// ---- POUs/System/Functions/FindINTFieldFragmented.TcPOU
FUNCTION FindINTFieldFragmented : INT
VAR_INPUT
    FieldName : STRING(254);
    Str1 : STRING(254);
    Str2 : STRING(254);
END_VAR
VAR_OUTPUT
    Valid : BOOL;
END_VAR
VAR
    value : DINT;
END_VAR

FindINTFieldFragmented := -9999;
value := FindDINTFieldFragmented(FieldName := FieldName, Str1 := Str1, Str2 := Str2, Valid => Valid);
IF NOT Valid THEN RETURN; END_IF;
Valid := (value >= -32768) AND (value <= 32767);
IF Valid THEN FindINTFieldFragmented := DINT_TO_INT(value); END_IF;

END_FUNCTION

// ---- POUs/System/Functions/RemovePlusSign.TcPOU
FUNCTION RemovePlusSign : STRING(254)
VAR_INPUT
    inString : STRING(254);
END_VAR

// Preserve the reference behavior: remove only one leading plus sign.
RemovePlusSign := inString;
IF LEFT(inString, 1) = '+' THEN
    RemovePlusSign := RIGHT(inString, LEN(inString) - 1);
END_IF;

END_FUNCTION

// ---- POUs/System/Tests/FC_TestTIAFoundation.TcPOU
FUNCTION FC_TestTIAFoundation : DWORD
VAR
    value : WORD;
    success : BOOL;
    decoded : ID_Decoded_DUT;
    lamps : Stack_Lights_FB;
    result : STRING(254);
END_VAR

// Offline utility checks: return DWORD#0 when all checks pass.
// Invoke manually in an isolated test PLC. No physical I/O or global data is used.
// Failure bits identify the numbered checks below; no task call is installed.
FC_TestTIAFoundation := DWORD#0;

// Bit 0: set the highest WORD bit and preserve other bits.
value := WORD#16#0001;
success := Set_Bit_F(BIT_Number := 15, Bit_Value := TRUE, Variavel := value);
IF NOT success OR (value <> WORD#16#8001) THEN
    FC_TestTIAFoundation := FC_TestTIAFoundation OR DWORD#16#0001;
END_IF;
// Bit 1: FALSE is intentionally a no-op, not a reset operation.
success := Set_Bit_F(BIT_Number := 15, Bit_Value := FALSE, Variavel := value);
IF NOT success OR (value <> WORD#16#8001) THEN
    FC_TestTIAFoundation := FC_TestTIAFoundation OR DWORD#16#0002;
END_IF;
// Bit 2: reject out-of-range shifts without modifying the word.
success := Set_Bit_F(BIT_Number := 16, Bit_Value := TRUE, Variavel := value);
IF success OR (value <> WORD#16#8001) THEN
    FC_TestTIAFoundation := FC_TestTIAFoundation OR DWORD#16#0004;
END_IF;
// Bit 3: decimal ID decomposition.
success := ID_Decode_F(ID := 123456, ID_Decoded := decoded);
IF NOT success OR (decoded.Device_Type <> 12) OR
   (decoded.Level <> 34) OR (decoded.VTD <> 56) THEN
    FC_TestTIAFoundation := FC_TestTIAFoundation OR DWORD#16#0008;
END_IF;
// Bit 4: invalid ID must not retain the preceding decoded result.
success := ID_Decode_F(ID := -1, ID_Decoded := decoded);
IF success OR (decoded.Device_Type <> 0) OR (decoded.Level <> 0) OR (decoded.VTD <> 0) THEN
    FC_TestTIAFoundation := FC_TestTIAFoundation OR DWORD#16#0010;
END_IF;
// Bit 5: accept leading zero fields and the unassigned ID.
success := ID_Decode_F(ID := 0, ID_Decoded := decoded);
IF NOT success OR (decoded.Device_Type <> 0) OR (decoded.Level <> 0) OR (decoded.VTD <> 0) THEN
    FC_TestTIAFoundation := FC_TestTIAFoundation OR DWORD#16#0020;
END_IF;
// Bit 6: source-compatible SICK field spacing.
result := FindStringField(FieldName := 'Code', JsonStr := '{"Number" :"2", "Code" :"ABC123"}');
IF result <> 'ABC123' THEN
    FC_TestTIAFoundation := FC_TestTIAFoundation OR DWORD#16#0040;
END_IF;
// Bit 7: a barcode longer than the source's 10-character search window.
result := FindStringField(FieldName := 'Code', JsonStr := '{"Code":"123456789012345678901234567890"}');
IF result <> '123456789012345678901234567890' THEN
    FC_TestTIAFoundation := FC_TestTIAFoundation OR DWORD#16#0080;
END_IF;
// Bit 8: missing field returns empty after a previous successful call.
result := FindStringField(FieldName := 'Code', JsonStr := '{"Number":"3"}');
IF result <> '' THEN
    FC_TestTIAFoundation := FC_TestTIAFoundation OR DWORD#16#0100;
END_IF;
// Bit 9: an unterminated value must not be accepted.
result := FindStringField(FieldName := 'Code', JsonStr := '{"Code":"ABC');
IF result <> '' THEN
    FC_TestTIAFoundation := FC_TestTIAFoundation OR DWORD#16#0200;
END_IF;
// Bit 10: fault takes priority over automatic mode.
lamps(System_Auto := TRUE, Fault := TRUE, i_bFlash_05Hz := TRUE);
IF NOT lamps.Red OR lamps.Green OR lamps.Orange OR lamps.Yellow THEN
    FC_TestTIAFoundation := FC_TestTIAFoundation OR DWORD#16#0400;
END_IF;
// Bit 11: manual mode uses yellow/orange and clears red/green.
lamps(System_Auto := FALSE, Fault := FALSE, i_bFlash_05Hz := FALSE);
IF lamps.Red OR lamps.Green OR NOT lamps.Orange OR NOT lamps.Yellow THEN
    FC_TestTIAFoundation := FC_TestTIAFoundation OR DWORD#16#0800;
END_IF;
// Bit 12: upper ID boundary validation.
success := ID_Decode_F(ID := 1000000, ID_Decoded := decoded);
IF success OR (decoded.Device_Type <> 0) OR (decoded.Level <> 0) OR (decoded.VTD <> 0) THEN
    FC_TestTIAFoundation := FC_TestTIAFoundation OR DWORD#16#1000;
END_IF;

END_FUNCTION

// ---- POUs/System/Tests/FC_TestTIAParsing.TcPOU
FUNCTION FC_TestTIAParsing : DWORD
VAR
    valid : BOOL;
    booleanValue : BOOL;
    integerValue : INT;
    longValue : DINT;
    buffer : ARRAY[0..1024] OF BYTE;
    result : STRING(254);
    window1 : STRING(254);
    truncated : BOOL;
    i : INT;
END_VAR

// Run only in an isolated test PLC. Zero means all checks passed.
// Each set bit identifies the corresponding assertion below.
FC_TestTIAParsing := DWORD#0;
IF RemovePlusSign('+42') <> '42' THEN FC_TestTIAParsing := FC_TestTIAParsing OR SHL(DWORD#1, 0); END_IF;
IF RemovePlusSign('4+2') <> '4+2' THEN FC_TestTIAParsing := FC_TestTIAParsing OR SHL(DWORD#1, 1); END_IF;
booleanValue := FindBoolField(FieldName := 'x', JsonStr := '{"x": false, "y": true}', Valid => valid);
IF booleanValue OR NOT valid THEN FC_TestTIAParsing := FC_TestTIAParsing OR SHL(DWORD#1, 2); END_IF;
booleanValue := FindBoolField(FieldName := 'x', JsonStr := '{"y":true}', Valid => valid);
IF booleanValue OR valid THEN FC_TestTIAParsing := FC_TestTIAParsing OR SHL(DWORD#1, 3); END_IF;
booleanValue := FindBoolField(FieldName := 'x', JsonStr := '{"x" :$T true$R$N}', Valid => valid);
IF NOT booleanValue OR NOT valid THEN FC_TestTIAParsing := FC_TestTIAParsing OR SHL(DWORD#1, 4); END_IF;
integerValue := FindIntField(FieldName := 'x', JsonStr := '{"x":32767}', Valid => valid);
IF NOT valid OR (integerValue <> 32767) THEN FC_TestTIAParsing := FC_TestTIAParsing OR SHL(DWORD#1, 5); END_IF;
integerValue := FindIntField(FieldName := 'x', JsonStr := '{"x":-32768}', Valid => valid);
IF NOT valid OR (integerValue <> -32768) THEN FC_TestTIAParsing := FC_TestTIAParsing OR SHL(DWORD#1, 6); END_IF;
integerValue := FindIntField(FieldName := 'x', JsonStr := '{"x":32768}', Valid => valid);
IF valid OR (integerValue <> -9999) THEN FC_TestTIAParsing := FC_TestTIAParsing OR SHL(DWORD#1, 7); END_IF;
longValue := FindDINTFieldFragmented(FieldName := 'x', Str1 := '{"x":2147483647}', Str2 := '', Valid => valid);
IF NOT valid OR (longValue <> DINT#2147483647) THEN FC_TestTIAParsing := FC_TestTIAParsing OR SHL(DWORD#1, 8); END_IF;
longValue := FindDINTFieldFragmented(FieldName := 'x', Str1 := '{"x":-2147483648}', Str2 := '', Valid => valid);
IF NOT valid OR (longValue <> DINT#-2147483648) THEN FC_TestTIAParsing := FC_TestTIAParsing OR SHL(DWORD#1, 9); END_IF;
longValue := FindDINTFieldFragmented(FieldName := 'x', Str1 := '{"x":2147483648}', Str2 := '', Valid => valid);
IF valid OR (longValue <> -9999) THEN FC_TestTIAParsing := FC_TestTIAParsing OR SHL(DWORD#1, 10); END_IF;
integerValue := FindIntField(FieldName := 'x', JsonStr := '{"x":12.3}', Valid => valid);
IF valid THEN FC_TestTIAParsing := FC_TestTIAParsing OR SHL(DWORD#1, 11); END_IF;
integerValue := FindIntField(FieldName := 'x', JsonStr := '{"x":12', Valid => valid);
IF valid THEN FC_TestTIAParsing := FC_TestTIAParsing OR SHL(DWORD#1, 12); END_IF;
integerValue := FindIntField(FieldName := 'x', JsonStr := '{"x":-9999}', Valid => valid);
IF NOT valid OR (integerValue <> -9999) THEN FC_TestTIAParsing := FC_TestTIAParsing OR SHL(DWORD#1, 13); END_IF;
integerValue := FindINTFieldFragmented(FieldName := 'x', Str1 := 'partial', Str2 := ',"x":42}', Valid => valid);
IF NOT valid OR (integerValue <> 42) THEN FC_TestTIAParsing := FC_TestTIAParsing OR SHL(DWORD#1, 14); END_IF;
integerValue := FindINTFieldFragmented(FieldName := 'x', Str1 := '{"x":4', Str2 := '2}', Valid => valid);
IF valid THEN FC_TestTIAParsing := FC_TestTIAParsing OR SHL(DWORD#1, 15); END_IF;
FOR i := 0 TO 1024 DO buffer[i] := 0; END_FOR;
buffer[0] := 65; buffer[1] := 13; buffer[2] := 10; buffer[3] := 66;
result := ByteArrayToString(Lenght := 4, ByteArray := buffer, Truncated => truncated);
IF (result <> 'AB') OR truncated THEN FC_TestTIAParsing := FC_TestTIAParsing OR SHL(DWORD#1, 16); END_IF;
result := ByteArrayToString(Lenght := -1, ByteArray := buffer, Truncated => truncated);
IF (result <> '') OR NOT truncated THEN FC_TestTIAParsing := FC_TestTIAParsing OR SHL(DWORD#1, 17); END_IF;
FOR i := 0 TO 254 DO buffer[i] := 65; END_FOR;
result := ByteArrayToString(Lenght := 255, ByteArray := buffer, ByteArrayToString_1 => window1, Truncated => truncated);
IF (LEN(result) <> 254) OR (LEN(window1) <> 155) OR NOT truncated THEN FC_TestTIAParsing := FC_TestTIAParsing OR SHL(DWORD#1, 18); END_IF;
integerValue := FindIntField(FieldName := 'x', JsonStr := '{"x":01}', Valid => valid);
IF valid THEN FC_TestTIAParsing := FC_TestTIAParsing OR SHL(DWORD#1, 19); END_IF;

END_FUNCTION

// ---- POUs/VTD/Light_Bars_FB.TcPOU
FUNCTION_BLOCK Light_Bars_FB
VAR_INPUT
	VTD_Mode:  UINT;
	VTD_Speed:  INT;
	Fault:  BOOL;
	// Drive enable state of the VTD. Replaces the Siemens "SinaSpeed_VTD_DB_1".EnableAxis
	// (enable of the former G120 drive). Suggested source: VTD_Control.Motor.stStatus.bOutputStageEnabled (PI 1.2).
	i_bDriveEnabled:  BOOL;
END_VAR
VAR_OUTPUT
	Animation_B1:  BYTE;
	Color_B1:  BYTE;
	Speed_B1:  Byte;
	Animation_B2:  Byte;
	Color_B2:  Byte;
	Speed_B2:  BYTE;
END_VAR
VAR
END_VAR

//Commands for Light Bar

IF VTD_Mode = 0 AND NOT Fault THEN // (0)Disabled = No light  
    Animation_B1:= Animation_B2:= 0;
    
// SIEMENS-LEGACY: ELSIF VTD_Mode = 1 AND VTD_Speed = 0 AND  NOT Fault AND NOT "SinaSpeed_VTD_DB_1".EnableAxis THEN // (1)Manual= Yellow Stop
ELSIF VTD_Mode = 1 AND VTD_Speed = 0 AND  NOT Fault AND NOT i_bDriveEnabled THEN // (1)Manual= Yellow Stop
    Animation_B1 := Animation_B2 := 1;
    Color_B1 := Color_B2 := 4;
    
// SIEMENS-LEGACY: ELSIF VTD_Mode = 1 AND VTD_Speed > 0 AND VTD_Speed <= 33 AND  NOT Fault AND "SinaSpeed_VTD_DB_1".EnableAxis THEN // (1)Manual= Yellow until 33%
ELSIF VTD_Mode = 1 AND VTD_Speed > 0 AND VTD_Speed <= 33 AND  NOT Fault AND i_bDriveEnabled THEN // (1)Manual= Yellow until 33%
    Animation_B1 := Animation_B2 := 2;
    Speed_B1 := Speed_B2 := 2;
    Color_B1 := Color_B2 := 4;
    
ELSIF VTD_Mode = 1 AND VTD_Speed > 33 AND VTD_Speed <= 100 AND  NOT Fault THEN // (1)Manual= Yellow until 66%
    Animation_B1 := Animation_B2 := 2;
    Speed_B1 := Speed_B2 := 0;
    Color_B1 := Color_B2 := 4;
    
// ELSIF VTD_Mode = 1 AND VTD_Speed > 66 AND VTD_Speed <= 100 AND  NOT Fault THEN // (1)Manual= Yellow until 100%
//     Animation_B1 := Animation_B2 := 2;
//     Speed_B1 := Speed_B2 := 1;
//     Color_B1 := Color_B2 := 4;
    
// SIEMENS-LEGACY: ELSIF VTD_Mode = 2 AND VTD_Speed = 0 AND  NOT Fault AND NOT "SinaSpeed_VTD_DB_1".EnableAxis THEN // (2)Semi-auto = Blue Stop
ELSIF VTD_Mode = 2 AND VTD_Speed = 0 AND  NOT Fault AND NOT i_bDriveEnabled THEN // (2)Semi-auto = Blue Stop
    Animation_B1 := Animation_B2 := 1;
    Color_B1 := Color_B2 := 9;
    Speed_B1 := Speed_B2 := 0;
    
// SIEMENS-LEGACY: ELSIF VTD_Mode = 2 AND VTD_Speed > 0 AND VTD_Speed <= 33 AND  NOT Fault AND "SinaSpeed_VTD_DB_1".EnableAxis THEN // (2)Semi-auto = Blue until 33%
ELSIF VTD_Mode = 2 AND VTD_Speed > 0 AND VTD_Speed <= 33 AND  NOT Fault AND i_bDriveEnabled THEN // (2)Semi-auto = Blue until 33%
    Animation_B1 := Animation_B2 := 2;
    Speed_B1 := Speed_B2 := 2;
    Color_B1 := Color_B2 := 9;
    
ELSIF VTD_Mode = 2 AND VTD_Speed > 33 AND VTD_Speed <= 100 AND  NOT Fault THEN // (2)Semi-auto = Blue until 66%
    Animation_B1 := Animation_B2 := 2;
    Speed_B1 := Speed_B2 := 0;
    Color_B1 := Color_B2 := 9;
    
// ELSIF VTD_Mode = 2 AND VTD_Speed > 66 AND VTD_Speed <= 100 AND  NOT Fault THEN // (2)Semi-auto = Blue until 100%
//     Animation_B1 := Animation_B2 := 2;
//     Speed_B1 := Speed_B2 := 1;
//     Color_B1 := Color_B2 := 9;
    
// SIEMENS-LEGACY: ELSIF VTD_Mode = 3 AND VTD_Speed = 0 AND  NOT Fault AND NOT "SinaSpeed_VTD_DB_1".EnableAxis THEN // (3)Auto = Green Stop
ELSIF VTD_Mode = 3 AND VTD_Speed = 0 AND  NOT Fault AND NOT i_bDriveEnabled THEN // (3)Auto = Green Stop
    Animation_B1 := Animation_B2 := 1;
    Color_B1 := Color_B2 := 0;
    
// SIEMENS-LEGACY: ELSIF VTD_Mode = 3 AND VTD_Speed > 0 AND VTD_Speed <= 33 AND  NOT Fault AND "SinaSpeed_VTD_DB_1".EnableAxis THEN // (3)Auto = Green until 33%
ELSIF VTD_Mode = 3 AND VTD_Speed > 0 AND VTD_Speed <= 33 AND  NOT Fault AND i_bDriveEnabled THEN // (3)Auto = Green until 33%
    Animation_B1 := Animation_B2 := 2;
    Speed_B1 := Speed_B2 := 2;
    Color_B1 := Color_B2 := 0;
    
ELSIF VTD_Mode = 3 AND VTD_Speed > 33 AND VTD_Speed <= 100 AND  NOT Fault THEN // (3)Auto = Green until 66%
    Animation_B1 := Animation_B2 := 2;
    Speed_B1 := Speed_B2 := 0;
    Color_B1 := Color_B2 := 0;
    
// ELSIF VTD_Mode = 3 AND VTD_Speed > 66 AND VTD_Speed <= 100 AND  NOT Fault THEN // (3)Auto = Green until 100%
//     Animation_B1 := Animation_B2 := 2;
//     Speed_B1 := Speed_B2 := 1;
//     Color_B1 := Color_B2 := 0;
    
ELSIF VTD_Mode = 4 AND VTD_Speed = 0 AND  NOT Fault THEN // (4)Tech = Orange Stop
    Animation_B1 := Animation_B2 := 1;
    Color_B1 := Color_B2 := 2;
    
ELSIF VTD_Mode = 4 AND VTD_Speed > 0 AND VTD_Speed <= 33 AND  NOT Fault THEN // (4)Tech = Orange until 33%
    Animation_B1 := Animation_B2 := 2;
    Speed_B1 := Speed_B2 := 2;
    Color_B1 := Color_B2 := 2;
    
ELSIF VTD_Mode = 4 AND VTD_Speed > 33 AND VTD_Speed <= 66 AND  NOT Fault THEN // (4)Tech = Orange until 66%
    Animation_B1 := Animation_B2 := 2;
    Speed_B1 := Speed_B2 := 0;
    Color_B1 := Color_B2 := 2;
    
ELSIF VTD_Mode = 4 AND VTD_Speed > 66 AND VTD_Speed <= 100 AND  NOT Fault THEN // (4)Tech = Orange until 100%
    Animation_B1 := Animation_B2 := 2;
    Speed_B1 := Speed_B2 := 1;
    Color_B1 := Color_B2 := 2;
    
ELSIF VTD_Mode = 5 AND VTD_Speed = 0 AND  NOT Fault THEN // (5)Maintenance = White Stop
    Animation_B1 := Animation_B2 := 1;
    Color_B1 := Color_B2 := 19;
    
ELSIF VTD_Mode = 5 AND VTD_Speed > 0 AND VTD_Speed <= 33 AND  NOT Fault THEN // (5)Maintenance = White until 33%
    Animation_B1 := Animation_B2 := 2;
    Speed_B1 := Speed_B2 := 2;
    Color_B1 := Color_B2 := 19;
    
ELSIF VTD_Mode = 5 AND VTD_Speed > 33 AND VTD_Speed <= 66 AND  NOT Fault THEN // (5)Maintenance = White until 66%
    Animation_B1 := Animation_B2 := 2;
    Speed_B1 := Speed_B2 := 0;
    Color_B1 := Color_B2 := 19;
    
ELSIF VTD_Mode = 5 AND VTD_Speed > 66 AND VTD_Speed <= 100 AND  NOT Fault THEN // (5)Maintenance = White until 100%
    Animation_B1 := Animation_B2 := 2;
    Speed_B1 := Speed_B2 := 1;
    Color_B1 := Color_B2 := 19;
    
ELSIF Fault THEN // Fault = Flash Red
    Animation_B1:= Animation_B2 := 2;
    Color_B1:=Color_B2 := 1;
END_IF;

END_FUNCTION_BLOCK

// ---- POUs/VTD/VTD_FB.TcPOU
FUNCTION_BLOCK VTD_FB
VAR_INPUT
	System_no:  UINT;
	Safety_OK:  BOOL;
	Cnv_Sensors:  Cnv_Inputs_DUT;
	VTD_Settings:  VTD_Settings_DUT;
	Bypass_DP:  BOOL;
// 	Bypass:  Safety_Bypass_RemotePanel;
END_VAR
VAR_OUTPUT
END_VAR
VAR_IN_OUT
	VTD_Control:  VTD_Control_DUT;
	LE_Bypass_HMI:  BOOL;
END_VAR
VAR
	State:  UINT;
	Last_State:  UINT;
	I_State:  UInt;
	LD_Timer_1:  TON;
	LD_Timer:  TON;
	DP_Timer:  TON;
	Watchdog:  TON;
	CS_TImer:  TON;
	Interlock_Timer:  TON;
	MainSetpoint:  Int;
	Position_Offset:  Real;
	ChangeToLow:  Array[1..4] of DInt;
	DestPosition:  Real;
	SetUpSpeed:  UInt;
	LevelBelowExtractor:  UInt;
	IEC_Timer_0_Instance:  TON;
	DestinationLevel:  UInt;
	CurrentlLevel:  UInt;
	VTD_ID_Decoded:  ID_Decoded_DUT;
	Cnv_ID_Decoded:  ARRAY[1..2] OF ID_Decoded_DUT;
	IEC_Timer_0_Instance_1:  TON;
	IEC_Timer_0_Instance_2:  TON;
	VTD_ControlInstructionTask_ID_Old:  Int;
	R_Execulte:  R_TRIG;
	R_AutomatcMode:  R_TRIG;
	T_Encoders_Difference:  TON;
	T_LE_Error:  TON;
	T_Setpoint_Delay:  TON;
	Distance_mm:  Real;
	TravelTime_s:  UInt;
	LE_Prev_mm:  Real;
	DeltaPos_mm:  Real;
	SampleTime_s:  Real;
	VTDSpeed_mm_s:  Real;
	T_Speed:  TON;
	Speed_mm_per_percent:  Real;
	Speed_mm_s:  Real;
	TravelTime_ms:  UInt;
	Watchdog_PT:  Time;
	Position_OLD:  Real;
	R_Position_OLD:  R_TRIG;

	// VTD drive: SEW MOVIPRO, MOVIKIT Positioning Drive (region "VFD")
	fbSewDrive:  FB_SEW_Drive;
	bDriveMoveRequest:  BOOL;
	bDriveEnable:  BOOL;
	bDriveFaultReset:  BOOL;
	rSpeedSetpoint:  REAL;              // [user units], signed
	rAccelerationFactor_pct:  REAL;     // [%] of SEW_Ramp_At_100pct
	uiDriveRamp:  UINT;                 // [user units]
	diPalletWeight:  DINT;
END_VAR

VAR_TEMP
	Level_Accuracy:  STRING;
	i:  UINT;
	Upper_limit:  Bool;
	Ultimate_SlowDown:  Bool;
	Ultimate_Creep:  Bool;
	Lower_Limit:  Bool;
	Level_Detect:  Bool;
	Level_Detect1:  Bool;
	Level_Detect2:  Bool;
	DP2_Extended:  Bool;
	DP2_Retracted:  Bool;
	DP1_Extended:  Bool;
	DP1_Retracted:  Bool;
	Chain_Slack_1:  Bool;
	Chain_Slack_2:  Bool;
	Chain_Slack_3:  Bool;
	Chain_Slack_4:  Bool;
	DP1_Retract:  Bool;
	DP1_Extend:  Bool;
	DP2_Retract:  Bool;
	DP2_Extend:  Bool;
	Cnvs1_NotExtended:  Bool;
	Cnvs2_NotExtended:  Bool;
	Stoppers_NotExtended:  Bool;
	MainSetpoint1:  Int;
	HMI_Reset:  BOOL;
END_VAR

// //Execute
// R_Execulte(CLK := VTD_Control.Instruction.Execulte);
// 
// IF VTD_Control.Mode = 3 THEN
//     VTD_Control.Instruction.Enable := TRUE;
// END_IF;
// 
// VTD_Control.Enabled := VTD_Control.Instruction.Enable;
// 
// VTD_Control.Mode := VTD_Control.Instruction.Mode_Change;
// 
// IF NOT VTD_Control.Enabled AND NOT VTD_Control.Error THEN
//     State := 0;
// END_IF;
// 
// //MANUAL MODE
// IF (VTD_Control.Mode = 1 OR VTD_Control.Mode = 5) AND NOT VTD_Control.Error AND VTD_Control.Enabled THEN
//     State := 500;
// END_IF;
// 
// (*
// TODO:
// 
// Mode select is done via the HMI. Might add external mode select switches.
//         
//         Mode select mask:
//         0: Disabled
//         1: Manual
//         2: Semi-Auto
//         3: Auto
//         4: Teach
//         5: Maintenance
//         
// Device ID Format: XXYYZZ    
// XX = Device type   
//     01   VTD
//     10  Cnv_Front_of_VTD
//     11  Cnv_Rear_of_VTD
//     12  Cnv_On_Extractor
//     20  Safety_Stop_Front_of_VTD
//     21  Safety_Stop_Rear_of_VTD
// YY = Floor   
// ZZ = VTD Connected to 
// *)
// 
// {region "Sensor allocations"}
//     //Assign inputs to local vars
//     Upper_limit := VTD_Control.Inputs.Upper_limit;
//     Ultimate_SlowDown := VTD_Control.Inputs.Ultimate_SlowDown;
//     Ultimate_Creep := VTD_Control.Inputs.Ultimate_Creep;
//     Lower_Limit := VTD_Control.Inputs.Lower_Limit;
//     Level_Detect1 := VTD_Control.Inputs.Level_Detect1;
//     Level_Detect2 := VTD_Control.Inputs.Level_Detect2;
//     DP1_Extended := VTD_Control.Inputs.DP1_Extended;
//     DP1_Retracted := VTD_Control.Inputs.DP1_Retracted;
//     DP2_Extended := VTD_Control.Inputs.DP2_Extended;
//     DP2_Retracted := VTD_Control.Inputs.DP2_Retracted;
//     Chain_Slack_1 := VTD_Control.Inputs.Chain_Slack_1;
//     Chain_Slack_2 := VTD_Control.Inputs.Chain_Slack_2;
//     Chain_Slack_3 := VTD_Control.Inputs.Chain_Slack_3;
//     Chain_Slack_4 := VTD_Control.Inputs.Chain_Slack_4;
//     VTD_Control.LinearEnc := VTD_Control.Inputs.LE_Position;
//     VTD_Control.AE := VTD_Control.Inputs.AE_Position_1;
// {endregion}
// 
// {region "Cyclic Checks"}
//     // Check for Pallet
//     IF Cnv_Sensors.Forward_Sensor OR Cnv_Sensors.Backward_Sensor THEN
//         VTD_Control.Pallet_Loaded := 1;//'Unknown';
//     ELSE
//         //No Pallet
//         VTD_Control.Pallet_Loaded := 0;//'None';
//     END_IF;
//     
//     //Docking pins
//         IF DP1_Extended AND DP2_Extended THEN
//             VTD_Control.LP_State := 1; //'Extended'
//         ELSIF DP1_Retracted AND DP2_Retracted THEN
//             VTD_Control.LP_State := 2; //'Retracted'
//         ELSE
//             VTD_Control.LP_State := 0; //'Unknown'
//         END_IF;
//         
//         VTD_Control.DP_Extended := VTD_Control.LP_State = 1;
//     
//     // Level detect
//     Level_Detect := Level_Detect1 AND Level_Detect2;
//     
//     //VTD extractor is docked
//     IF DP1_Extended AND DP2_Extended AND Level_Detect AND
//         (VTD_Control.LinearEnc - VTD_Settings.Teach_Values.Levels_LE[LevelBelowExtractor]) <= VTD_Settings.Level_Detect_LE THEN
//         VTD_Control.Docked := TRUE;
//     ELSE
//         VTD_Control.Docked := FALSE;
//     END_IF;
//     
//     //Ultimate stop checks
//     IF (VTD_Control.LinearEnc < VTD_Settings.Slowdown_Count_LE OR VTD_Control.LinearEnc > VTD_Settings.Teach_Values.Levels_LE[VTD_Settings.Highest_Level] - VTD_Settings.Slowdown_Count_LE) AND
//         Ultimate_Creep AND Ultimate_SlowDown AND VTD_Control.Running THEN
//         VTD_Control.Motor_Speed := VTD_Settings.Creep_Speed;
//         VTD_Control.Warning := 3; // Overtravel creep zone reached
//     ELSIF (VTD_Control.LinearEnc < VTD_Settings.Slowdown_Count_LE OR VTD_Control.LinearEnc > VTD_Settings.Teach_Values.Levels_LE[VTD_Settings.Highest_Level] - VTD_Settings.Slowdown_Count_LE) AND
//         NOT Ultimate_Creep AND Ultimate_SlowDown AND VTD_Control.Running THEN
//         VTD_Control.Motor_Speed := VTD_Settings.Slow_Speed; // Overtravel slow zone reached
//     END_IF;
//     
//     //Update Variables
//     IF VTD_Control.Current_Task_Type = 0 OR VTD_Control.Current_Task_Type = 1 THEN
//         VTD_Control.SM_State := State;
//     ELSIF VTD_Control.Current_Task_Type = 2 OR VTD_Control.Current_Task_Type = 3 THEN
//         VTD_Control.SM_State := I_State;
//     END_IF;
//     
//     FOR i := VTD_Settings.Lowest_Level TO VTD_Settings.Highest_Level DO
//         IF NOT Control.LCnv_Sys[System_no].Cnv_Level[i].Cnv1.Safety_Stop_Cnrl.Inputs.DP_Extended THEN
//             Cnvs1_NotExtended := true;
//         END_IF;
//         IF NOT Control.LCnv_Sys[System_no].Cnv_Level[i].Cnv2.Safety_Stop_Cnrl.Inputs.DP_Extended THEN
//             Cnvs2_NotExtended := true;
//         END_IF;
//     END_FOR;
//     
//     //Confirm whish level is below the extractor
//     FOR i := VTD_Settings.Lowest_Level TO VTD_Settings.Highest_Level DO
//         IF VTD_Control.LinearEnc >= (VTD_Settings.Teach_Values.Levels_LE[i] - VTD_Settings.Level_Detect_LE) THEN
//             LevelBelowExtractor := i;
//         END_IF;
//     END_FOR;
//     
//     Stoppers_NotExtended := Cnvs1_NotExtended (*AND Cnvs2_NotExtended*);
//     
//     //AE ERROR
//     IF VTD_Control.Inputs.AE_Status_2.15 THEN
//         VTD_Control.AE_Error := 1;
//     ELSE
//         VTD_Control.AE_Error := 0;
//     END_IF;
//     
//     //Encoder Delta
//     VTD_Control.Encoder_Delta := ABS(VTD_Control.AE - VTD_Control.LinearEnc);
//     
//     //CURRENT LEVEL
//     FOR i := VTD_Settings.Lowest_Level TO VTD_Settings.Highest_Level DO
//         IF ABS(VTD_Control.LinearEnc - VTD_Settings.Teach_Values.Levels_LE[i]) <= VTD_Settings.VTD_Level_Granularity AND Level_Detect THEN
//             VTD_Control.Current_Level := i;
//             EXIT;
//         ELSE
//             VTD_Control.Current_Level := 0;
//         END_IF;
//     END_FOR;
//     
//     //SPEED mm/S
//     T_Speed(IN := TRUE,
//              PT := T#100MS);
//     
//     IF T_Speed.Q THEN
//         DeltaPos_mm := ABS(VTD_Control.LinearEnc - LE_Prev_mm);
//         VTDSpeed_mm_s := DeltaPos_mm / SampleTime_s;
//         LE_Prev_mm := VTD_Control.LinearEnc;
//         T_Speed(IN := FALSE,
//                  PT := T#0MS);
//     END_IF;
// {endregion}
// 
// {region "Auto/Semi-Auto Mode"}
//     CASE State OF
//         0: //Idle
//             Last_State := State;
//             VTD_Control.Motor_UP := FALSE;
//             VTD_Control.Motor_Down := FALSE;
//             VTD_Control.Motor_Speed := 0; // SEW: was Motor.Speed
//             DestinationLevel := CurrentlLevel := 0;
//             VTD_Control.Stopped := TRUE;
//             Watchdog(IN := FALSE,
//                           PT := T#0S);
//             IF VTD_Control.Mode = 3 OR VTD_Control.Mode = 2 THEN
//                 IF VTD_Control.Instruction.Enable AND NOT VTD_Control.Error THEN
//                     State := 10;
//                 END_IF;
//             END_IF;
//             
//         10: //Standby
//             Last_State := State;
//             IF VTD_Control.Enabled AND NOT VTD_Control.Running AND VTD_Control.Instruction.Move_To_Level >= VTD_Settings.Lowest_Level AND
//                 VTD_Control.Instruction.Move_To_Level <= VTD_Settings.Highest_Level AND VTD_Control.Pallet_Loaded <> 1 AND
//                 ((VTD_Control.Instruction.Task_ID > 0 OR VTD_Control.Instruction.Task_Metadata <> '' AND VTD_Control.Mode = 3 AND Control.VTD_Order_Table[System_no].Task_Type = 1) OR
//                 (VTD_Control.Mode = 2 (*AND R_Execulte.Q*)))
//             THEN
//                 IF VTD_Control.Instruction.Move_To_Level = VTD_Control.Current_Level AND VTD_Control.Instruction.Move_To_Level <> 0 THEN
//                     VTD_Control.Warning := 1; //VTD already at level requested
//                     VTD_Control.Instruction.Move_To_Level := 0;
//                     //Go straght to the travel complete feedabck 
//                 ELSIF ((VTD_Control.Shuttle_Loaded = 0 OR VTD_Control.Shuttle_Loaded = 1) AND System_no <= 3)
//                     OR System_no > 3
//                 THEN //EVERYTHING OK
//                     DestinationLevel := VTD_Control.Instruction.Move_To_Level;
//                     CurrentlLevel := VTD_Control.Current_Level;
//                     VTD_Control.Current_Task_ID := VTD_Control.Instruction.Task_ID;
//                     VTD_Control.Running := TRUE;
//                     State := 20;
//                 END_IF;
//             END_IF;
// 
//         20: //Extend all safety stoppers that are not in the up position
//             Last_State := State;
//             VTD_Control.Done := FALSE;// To report to order table
//             FOR i := VTD_Settings.Lowest_Level TO VTD_Settings.Highest_Level DO
//                 IF NOT Control.LCnv_Sys[System_no].Cnv_Level[i].Cnv1.Safety_Stop_Cnrl.Inputs.DP_Extended THEN
//                     Control.LCnv_Sys[System_no].Cnv_Level[i].Cnv1.Safety_Stop_Cnrl.Instruction.Extend := TRUE;
//                 END_IF;
//                 IF NOT Control.LCnv_Sys[System_no].Cnv_Level[i].Cnv2.Safety_Stop_Cnrl.Inputs.DP_Extended THEN
//                     Control.LCnv_Sys[System_no].Cnv_Level[i].Cnv2.Safety_Stop_Cnrl.Instruction.Extend := TRUE;
//                 END_IF;
//             END_FOR;
//             State := 25;
//             
//         25: //Check to ensure the Safety stoppers are in the up position.
//             Last_State := State;
//             FOR i := VTD_Settings.Lowest_Level TO VTD_Settings.Highest_Level DO
//                 IF Control.LCnv_Sys[System_no].Cnv_Level[i].Cnv1.Safety_Stop_Cnrl.Inputs.DP_Extended THEN
//                     Control.LCnv_Sys[System_no].Cnv_Level[i].Cnv1.Safety_Stop_Cnrl.Instruction.Extend := FALSE;
//                 END_IF;
//                 IF Control.LCnv_Sys[System_no].Cnv_Level[i].Cnv2.Safety_Stop_Cnrl.Inputs.DP_Extended THEN
//                     Control.LCnv_Sys[System_no].Cnv_Level[i].Cnv2.Safety_Stop_Cnrl.Instruction.Extend := FALSE;
//                 END_IF;
//             END_FOR;
//             
//             IF Control.LCnv_Sys[System_no].Cnv_Level[2].Cnv1.Safety_Stop_Cnrl.Inputs.DP_Extended AND
//                 Control.LCnv_Sys[System_no].Cnv_Level[3].Cnv1.Safety_Stop_Cnrl.Inputs.DP_Extended AND
//                 Control.LCnv_Sys[System_no].Cnv_Level[4].Cnv1.Safety_Stop_Cnrl.Inputs.DP_Extended AND
//                 Control.LCnv_Sys[System_no].Cnv_Level[5].Cnv1.Safety_Stop_Cnrl.Inputs.DP_Extended AND
//                 Control.LCnv_Sys[System_no].Cnv_Level[6].Cnv1.Safety_Stop_Cnrl.Inputs.DP_Extended AND
//                 Control.LCnv_Sys[System_no].Cnv_Level[2].Cnv2.Safety_Stop_Cnrl.Inputs.DP_Extended AND
//                 Control.LCnv_Sys[System_no].Cnv_Level[3].Cnv2.Safety_Stop_Cnrl.Inputs.DP_Extended AND
//                 Control.LCnv_Sys[System_no].Cnv_Level[4].Cnv2.Safety_Stop_Cnrl.Inputs.DP_Extended AND
//                 Control.LCnv_Sys[System_no].Cnv_Level[5].Cnv2.Safety_Stop_Cnrl.Inputs.DP_Extended AND
//                 Control.LCnv_Sys[System_no].Cnv_Level[6].Cnv2.Safety_Stop_Cnrl.Inputs.DP_Extended
//             THEN
//                 State := 30;
//             END_IF;
//             
//         30: //Undock the VTD
//             Last_State := State;
//             IF LevelBelowExtractor >= VTD_Settings.Lowest_Level AND LevelBelowExtractor < VTD_Settings.Highest_Level THEN
//                 IF VTD_Control.Docked OR
//                     (VTD_Control.LinearEnc < VTD_Settings.Teach_Values.Levels_LE[LevelBelowExtractor] + 50) OR
//                     (VTD_Control.LinearEnc < VTD_Settings.Teach_Values.Levels_LE[LevelBelowExtractor + 1] AND
//                     VTD_Control.LinearEnc > VTD_Settings.Teach_Values.Levels_LE[LevelBelowExtractor + 1] - 10) THEN
//                     IF VTD_Control.LP_State = 1 THEN //extended
//                         VTD_Control.Motor_Speed := VTD_Settings.Dock_speed;
//                         VTD_Control.Motor_UP := TRUE;
//                         Position_Offset := VTD_Control.LinearEnc + 40;
//                         State := 35;
//                     ELSIF VTD_Control.LP_State = 2 THEN //retracted
//                         State := 45;
//                     ELSE //24:4 Docking pins in an known state
//                         Set_Bit_F(Bit_Number := 5,
//                                     Bit_Value := 1,
//                                     Variavel := VTD_Control.VTD_Errors.Error_Word_2);
//                     END_IF;
//                 ELSE
//                     Position_Offset := VTD_Control.LinearEnc - 5;
//                     State := 35;
//                 END_IF;
//             ELSIF LevelBelowExtractor = VTD_Settings.Highest_Level THEN
//                 IF VTD_Control.Docked OR
//                     (VTD_Control.LinearEnc < VTD_Settings.Teach_Values.Levels_LE[LevelBelowExtractor] + 50) THEN
//                     IF VTD_Control.LP_State = 1 THEN //extended
//                         VTD_Control.Motor_Speed := VTD_Settings.Dock_speed;
//                         VTD_Control.Motor_UP := TRUE;
//                         Position_Offset := VTD_Control.LinearEnc + 40;
//                         State := 35;
//                     ELSIF VTD_Control.LP_State = 2 THEN //retracted
//                         State := 45;
//                     ELSE //24:4 Docking pins in an known state
//                         Set_Bit_F(Bit_Number := 5,
//                                     Variavel := VTD_Control.VTD_Errors.Error_Word_2);
//                     END_IF;
//                 ELSE
//                     Position_Offset := VTD_Control.LinearEnc - 5;
//                     State := 35;
//                 END_IF;
//             END_IF;
//             
//         35: //Stop motor
//             Last_State := State;
//             IF NOT Level_Detect AND VTD_Control.LinearEnc >= Position_Offset THEN
//                 VTD_Control.Motor_Speed := 0;
//                 VTD_Control.Motor_UP := FALSE;
//                 State := 36;
//             END_IF;
//             
//         36: //Retract the docking pins
//             Last_State := State;
//                 DP2_Retract := DP1_Retract := TRUE;
//                 DP_Timer(IN := TRUE,
//                           PT := UINT_TO_TIME(VTD_Settings.Lockpins_Timeout_Retract));
//                 
//                 IF DP2_Retracted THEN
//                     DP2_Retract := FALSE;
//                 END_IF;
//                 IF VTD_Control.Inputs.DP1_Retracted THEN
//                     DP1_Retract := FALSE;
//                 END_IF;
//                 
//                 IF VTD_Control.LP_State = 2 THEN
//                     State := 40;
//                 END_IF;
//                 
//             40: //Check docking pins have been retracted
//                 Last_State := State;
//             IF VTD_Control.LP_State = 2 THEN
//                 DP_Timer(IN := FALSE,
//                           PT := T#0S);
//                 DP2_Retract := DP1_Retract := FALSE;
//                 State := 45;
//             END_IF;
//             
//         45: //Start moving towards the level required
//             Last_State := State;
//             //Check load type and set extractor speed
//             IF VTD_Control.Shuttle_Loaded = 0 AND VTD_Control.Pallet_Loaded = 0 THEN
//                 VTD_Control.Motor_Speed := VTD_Settings.Empty_Speed;
//             ELSIF VTD_Control.Shuttle_Loaded = 1 AND VTD_Control.Pallet_Loaded = 0 THEN
//                 VTD_Control.Motor_Speed := VTD_Settings.Shuttle_Speed;
//             ELSIF VTD_Control.Shuttle_Loaded = 0 AND (VTD_Control.Pallet_Loaded > 0) THEN
//                 VTD_Control.Motor_Speed := VTD_Settings.Pallet_Speed;
//             ELSIF VTD_Control.Shuttle_Loaded = 1 AND (VTD_Control.Pallet_Loaded > 0) THEN
//                 VTD_Control.Motor_Speed := VTD_Settings.Loaded_Speed;
//             END_IF;
//             
//             DestPosition := VTD_Settings.Teach_Values.Levels_LE[VTD_Control.Instruction.Move_To_Level];
//             SetUpSpeed := VTD_Control.Motor_Speed;
//             
//             // === DINAMIC WATCHDOG ===
//             Speed_mm_s := SetUpSpeed * Speed_mm_per_percent;
//             Distance_mm := ABS(DestPosition - VTD_Control.LinearEnc);
//             
//             //VTD needs to move up
//             IF VTD_Control.LinearEnc < DestPosition THEN
//                 VTD_Control.Motor_UP := TRUE;
//                 State := 50;
//                 //VTD needs to move down
//             ELSIF VTD_Control.LinearEnc > DestPosition THEN
//                 VTD_Control.Motor_Down := TRUE;
//                 State := 65; //change to 65
//             END_IF;
//             
//         50: //travel upwards to designated level
//             Last_State := State;
//             ChangeToLow[1] := ABS((VTD_Settings.Slowdown_Count_LE / 100) * 80); (* 80% *) //80  600mm
//             ChangeToLow[2] := ABS((VTD_Settings.Slowdown_Count_LE / 100) * 60); (* 60% *) //60
//             ChangeToLow[3] := ABS((VTD_Settings.Slowdown_Count_LE / 100) * 40); (* 40% *) //40
//             ChangeToLow[4] := ABS((VTD_Settings.Slowdown_Count_LE / 100) * 20); (* 20% *) //20 60
//             
//             //switch to fast freq Low UP
//             IF ABS(DestPosition - VTD_Control.LinearEnc) > VTD_Settings.Slowdown_Count_LE THEN
//                 VTD_Control.Motor_Speed := SetUpSpeed; //5
//                 //switch to low freq
//             ELSIF ABS(DestPosition - VTD_Control.LinearEnc) <= VTD_Settings.Slowdown_Count_LE
//                 AND ABS(DestPosition - VTD_Control.LinearEnc) > ChangeToLow[1] THEN
//                 VTD_Control.Motor_Speed := VTD_Settings.Slow_Calib_Speed * 1.8; //5 * 1.8 = 9%
//             ELSIF ABS(DestPosition - VTD_Control.LinearEnc) <= ChangeToLow[1]
//                 AND ABS(DestPosition - VTD_Control.LinearEnc) > ChangeToLow[2] THEN
//                 VTD_Control.Motor_Speed := VTD_Settings.Slow_Calib_Speed * 1.6; //5 * 1.6 = 8%
//             ELSIF ABS(DestPosition - VTD_Control.LinearEnc) <= ChangeToLow[2]
//                 AND ABS(DestPosition - VTD_Control.LinearEnc) > ChangeToLow[3] THEN
//                 VTD_Control.Motor_Speed := VTD_Settings.Slow_Calib_Speed * 1.4; //5 * 1.4 = 7%
//             ELSIF ABS(DestPosition - VTD_Control.LinearEnc) <= ChangeToLow[3]
//                 AND ABS(DestPosition - VTD_Control.LinearEnc) > ChangeToLow[4] THEN
//                 VTD_Control.Motor_Speed := VTD_Settings.Slow_Calib_Speed * 1.2; //5 * 1.2 = 6%
//             ELSIF ABS(DestPosition - VTD_Control.LinearEnc) <= ChangeToLow[4] THEN
//                 VTD_Control.Motor_Speed := VTD_Settings.Slow_Calib_Speed; //5%
//                 State := 55;
//             END_IF;
//             
//             // Timeout in ms
//             IF Speed_mm_s > 0 THEN
//                 TravelTime_ms := REAL_TO_UINT((Distance_mm / Speed_mm_s) * 1500.0);  // 1.5x safety factor
//                 IF TravelTime_ms < 5000 THEN
//                     TravelTime_ms := 5000; // mínimum 5s
//                 END_IF;
//             ELSE
//                 TravelTime_ms := 30000; // fallback 30s 
//             END_IF;
//             
//             Watchdog_PT := UINT_TO_TIME(TravelTime_ms);
//             
//             Watchdog.TON(IN := TRUE,
//                           PT := Watchdog_PT);
//             
//             
//         55: // Travel upwards using slow speed towards required floor
//             Last_State := State;
//             IF VTD_Control.LinearEnc > VTD_Settings.Teach_Values.Levels_LE[VTD_Control.Instruction.Move_To_Level] - VTD_Settings.Creep_Count_LE
//             THEN
//                 VTD_Control.Motor_Speed := VTD_Settings.Creep_Speed; //3% - 60mm 
//                 State := 60;
//             END_IF;
//             
//         60: // Travel past the level in order to extend the docking pins
//             Last_State := State;
//             IF VTD_Control.LinearEnc > VTD_Settings.Teach_Values.Levels_LE[VTD_Control.Instruction.Move_To_Level] + VTD_Settings.Creep_Count_LE
//             THEN
//                 VTD_Control.Motor_Speed := 0;
//                 VTD_Control.Motor_UP := FALSE;
//                 VTD_Control.Motor_Down := FALSE;
//                 State := 80;
//             END_IF;
//             
//         65: //travel Downwards to designated level   
//             Last_State := State;
//             ChangeToLow[1] := ABS((VTD_Settings.Slowdown_Count_LE / 100) * 80); (* 80% *) //80
//             ChangeToLow[2] := ABS((VTD_Settings.Slowdown_Count_LE / 100) * 60); (* 60% *) //60
//             ChangeToLow[3] := ABS((VTD_Settings.Slowdown_Count_LE / 100) * 40); (* 40% *) //40
//             ChangeToLow[4] := ABS((VTD_Settings.Slowdown_Count_LE / 100) * 20); (* 20% *) //20
//             //switch to fast freq Low UP
//             IF ABS(DestPosition - VTD_Control.LinearEnc) > VTD_Settings.Slowdown_Count_LE THEN
//                 VTD_Control.Motor_Speed := SetUpSpeed;
//                 //switch to low freq
//             ELSIF ABS(DestPosition - VTD_Control.LinearEnc) <= VTD_Settings.Slowdown_Count_LE
//                 AND ABS(DestPosition - VTD_Control.LinearEnc) > ChangeToLow[1] THEN
//                 VTD_Control.Motor_Speed := REAL_TO_UINT(VTD_Settings.Slow_Calib_Speed * 1.8);
//             ELSIF ABS(DestPosition - VTD_Control.LinearEnc) <= ChangeToLow[1]
//                 AND ABS(DestPosition - VTD_Control.LinearEnc) > ChangeToLow[2] THEN
//                 VTD_Control.Motor_Speed := REAL_TO_UINT(VTD_Settings.Slow_Calib_Speed * 1.6);
//             ELSIF ABS(DestPosition - VTD_Control.LinearEnc) <= ChangeToLow[2]
//                 AND ABS(DestPosition - VTD_Control.LinearEnc) > ChangeToLow[3] THEN
//                 VTD_Control.Motor_Speed := REAL_TO_UINT(VTD_Settings.Slow_Calib_Speed * 1.4);
//             ELSIF ABS(DestPosition - VTD_Control.LinearEnc) <= ChangeToLow[3]
//                 AND ABS(DestPosition - VTD_Control.LinearEnc) > ChangeToLow[4] THEN
//                 VTD_Control.Motor_Speed := REAL_TO_UINT(VTD_Settings.Slow_Calib_Speed * 1.2);
//             ELSIF ABS(DestPosition - VTD_Control.LinearEnc) <= ChangeToLow[4] THEN
//                 VTD_Control.Motor_Speed := VTD_Settings.Slow_Calib_Speed;
//                 State := 70;
//             END_IF;
//             
//             // Timeout in ms
//             IF Speed_mm_s > 0 THEN
//                 TravelTime_ms := REAL_TO_UINT((Distance_mm / Speed_mm_s) * 2000.0);  // 1.5x safety factor
//                 IF TravelTime_ms < 5000 THEN
//                     TravelTime_ms := 5000; // mínimum 5s
//                 END_IF;
//             ELSE
//                 TravelTime_ms := 30000; // fallback 30s 
//             END_IF;
//             
//             Watchdog_PT := UINT_TO_TIME(TravelTime_ms);
//             
//             Watchdog(IN := TRUE,
//                      PT := Watchdog_PT);
//             
//         70: // Travel downwards using slow speed towards required floor 
//             Last_State := State;
//             IF VTD_Control.LinearEnc < VTD_Settings.Teach_Values.Levels_LE[VTD_Control.Instruction.Move_To_Level] + VTD_Settings.Creep_Count_LE
//             THEN
//                 VTD_Control.Motor_Speed := 0;
//                 VTD_Control.Motor_UP := FALSE;
//                 VTD_Control.Motor_Down := FALSE;
//                 State := 80;
//             END_IF;
//             
//         80: //Extend Docking pins
//             Last_State := State;
//             IF VTD_Control.LP_State = 2 AND NOT Level_Detect THEN
//                 DP1_Extend := DP2_Extend := TRUE;
//                 DP_Timer(IN := TRUE,
//                           PT := UINT_TO_TIME(VTD_Settings.Lockpins_Timeout_Extend));
//             ELSIF VTD_Control.LP_State <> 1 AND NOT Level_Detect THEN
//                 DP1_Extend := DP2_Extend := TRUE;
//             ELSIF VTD_Control.LP_State = 1 THEN
//                 State := 85;
//             END_IF;
//             
//             
//         85: // Wait for docking pins to extend
//             Last_State := State;
//             IF VTD_Control.LP_State = 1 AND NOT Level_Detect THEN
//                 DP_Timer(IN := FALSE,
//                           PT := T#0S);
//                 DP1_Extend := DP2_Extend := FALSE;
//                 VTD_Control.Motor_Speed := VTD_Settings.Dock_speed;
//                 VTD_Control.Motor_Down := TRUE;
//                 State := 90;
//             END_IF;
//             
//         90: // Dock the VTD
//             Last_State := State;
//             //Using the LE for comparation and Release tension in the VTD chain
//             IF ABS(VTD_Control.LinearEnc - DestPosition) <= (VTD_Settings.Level_Detect_LE) AND NOT CS_TImer.Q THEN
//                 CS_TImer(IN := TRUE,
//                           PT := UINT_TO_TIME(VTD_Settings.Chain_Slack_Timeout));
//             END_IF;
//             IF CS_TImer.Q THEN
//                 VTD_Control.Motor_Speed := 0;
//                 VTD_Control.Motor_Down := FALSE;
//                 CS_TImer(IN := FALSE,
//                           PT := T#0S);
//                 State := 95;
//             END_IF;
//             
//         95: // Dock the VTD
//             Last_State := State;
//             //Check the level detect sensors
//             IF (Level_Detect1 AND NOT Level_Detect2) OR
//                 (NOT Level_Detect1 AND Level_Detect2) THEN
//                 LD_Timer(IN := TRUE,
//                           PT := UINT_TO_TIME(VTD_Settings.Level_Detect_Timeout));
//             ELSIF NOT Level_Detect1 AND NOT Level_Detect2 THEN
//                 LD_Timer_1(IN := TRUE,
//                             PT := UINT_TO_TIME(VTD_Settings.Level_Detect_Timeout * 5));
//             ELSE
//                 LD_Timer(IN := FALSE,
//                           PT := T#0S);
//                 LD_Timer_1(IN := FALSE,
//                             PT := T#0S);
//             END_IF;
//             
//             IF Level_Detect THEN
//                 Watchdog(IN := FALSE,
//                           PT := T#0S);
//                 State := 100;
//             END_IF;
//             
//         100: //Wait for Movement completion ack  
//             Last_State := State;
//             //Reset timers
//             VTD_Control.Instruction.Move_To_Level := 0;
//             DP_Timer(IN := FALSE,
//                       PT := T#0S);
//             Watchdog(IN := FALSE,
//                       PT := T#0S);
//             LD_Timer(IN := FALSE,
//                       PT := T#0S);
//             CS_TImer(IN := FALSE,
//                       PT := T#0S);
//             LD_Timer_1(IN := FALSE,
//                         PT := T#0S);
//             
//             VTD_Control.Motor_Speed := 0;
//             VTD_Control.Current_Task_ID := 0;
//             VTD_Control.Running := FALSE;
//             State := 0;
//             
//         400: // Error state
//             VTD_Control.Instruction.Move_To_Level := 0;
//             VTD_Control.Done := FALSE;// To report to order table
//             // SEW: Motor_UP/Motor_Down := FALSE removes enable/start in region "VFD"
//             VTD_Control.Motor_UP := FALSE;
//             VTD_Control.Motor_Down := FALSE;
//             VTD_Control.Running := FALSE;
//             VTD_Control.Stopped := TRUE;
//             VTD_Control.Motor_Speed := 0; // SEW: was Motor.Speed/Forward/Reverse
//             DP1_Extend := DP2_Extend := FALSE;
//             DP1_Retract := DP2_Retract := FALSE;
//             FOR i := VTD_Settings.Lowest_Level TO VTD_Settings.Highest_Level DO
//                 Control.LCnv_Sys[System_no].Cnv_Level[i].Cnv1.Safety_Stop_Cnrl.Instruction.Extend := FALSE;
//                 Control.LCnv_Sys[System_no].Cnv_Level[i].Cnv2.Safety_Stop_Cnrl.Instruction.Extend := FALSE;
//             END_FOR;
//             //Reset timers
//             DP_Timer(IN := FALSE,
//                       PT := T#0S);
//             Watchdog(IN := FALSE,
//                       PT := T#0S);
//             LD_Timer(IN := FALSE,
//                       PT := T#0S);
//             CS_TImer(IN := FALSE,
//                       PT := T#0S);
//             LD_Timer_1(IN := FALSE,
//                         PT := T#0S);
//             IF VTD_Control.Instruction.Reset OR Reset_All OR HMI_Reset THEN
//                 VTD_Control.Error := FALSE;
//                 VTD_Control.Warning := 0;
//                 VTD_Control.Stopped := FALSE;
//                 VTD_Control.Current_Task_Type := 0;
//                 VTD_Control.VTD_Errors.Error_Word_1 := 0;
//                 VTD_Control.VTD_Errors.Error_Word_2 := 0;
//                 VTD_Control.VTD_Errors.Error_Word_3 := 0;
//                 VTD_Control.VTD_Errors.Error_Word_4 := 0;
//                 VTD_Control.VTD_Errors.Error_Word_5 := 0;
//                 State := 0;
//             END_IF;
//             
//         500: //MANUAL MODE
//             IF VTD_Control.Error = 0 AND VTD_Control.Enabled THEN
//                 //VTD
//                 IF VTD_Control.Instruction.Manual_Up AND NOT Upper_limit THEN
//                     VTD_Control.Motor_UP := TRUE;
//                     VTD_Control.Stopped := FALSE;
//                     VTD_Control.Running := TRUE;
//                     IF NOT (Ultimate_SlowDown OR Ultimate_Creep) THEN
//                         VTD_Control.Motor_Speed := VTD_Settings.Manual_Speed;
//                     END_IF;
//                 ELSIF VTD_Control.Instruction.Manual_Down AND NOT Lower_Limit THEN
//                     VTD_Control.Motor_Down := TRUE;
//                     VTD_Control.Stopped := FALSE;
//                     VTD_Control.Running := TRUE;
//                     IF VTD_Control.LinearEnc <= VTD_Settings.Teach_Values.Levels_LE[LevelBelowExtractor] + 300 AND VTD_Control.LP_State = 1 THEN
//                         VTD_Control.Motor_Speed := VTD_Settings.Creep_Speed;
//                     ELSIF NOT (Ultimate_SlowDown OR Ultimate_Creep) THEN
//                         VTD_Control.Motor_Speed := VTD_Settings.Manual_Speed;
//                     END_IF;
//                 ELSE
//                     VTD_Control.Motor_Speed := 0;
//                     VTD_Control.Stopped := TRUE;
//                     VTD_Control.Running := FALSE;
//                     VTD_Control.Motor_Down := FALSE;
//                     VTD_Control.Motor_UP := FALSE;
//                 END_IF;
//                 
//                 //DOCKING PINS 2 
//                 IF NOT VTD_Control.Running AND VTD_Control.Instruction.Manual_LP_Extend
//                     AND NOT DP2_Extended THEN
//                     DP2_Extend := TRUE;
//                 ELSIF NOT VTD_Control.Running AND VTD_Control.Instruction.Manual_LP_Retract
//                     AND NOT DP2_Retracted THEN
//                     DP2_Retract := TRUE;
//                 ELSE
//                     DP2_Extend := FALSE;
//                     DP2_Retract := FALSE;
//                 END_IF;
//                 
//                 //DOCKING PINS 1 
//                 IF NOT VTD_Control.Running AND VTD_Control.Instruction.Manual_LP_Extend
//                     AND NOT DP1_Extended THEN
//                     DP1_Extend := TRUE;
//                 ELSIF NOT VTD_Control.Running AND VTD_Control.Instruction.Manual_LP_Retract
//                     AND NOT DP1_Retracted THEN
//                     DP1_Retract := TRUE;
//                 ELSE
//                     DP1_Extend := FALSE;
//                     DP1_Retract := FALSE;
//                 END_IF;
//                 
//                 IF VTD_Control.Mode <> 1 AND VTD_Control.Mode <> 5 THEN
//                     State := 0;
//                 END_IF;
//                 
//                 IF DP2_Extend OR DP1_Extend THEN
//                     DP_Timer(IN := TRUE,
//                               PT := UINT_TO_TIME(VTD_Settings.Lockpins_Timeout_Extend));
//                 ELSIF DP2_Retract OR DP1_Retract THEN
//                     DP_Timer(IN := TRUE,
//                               PT := UINT_TO_TIME(VTD_Settings.Lockpins_Timeout_Retract));
//                 ELSE
//                     DP_Timer(IN := FALSE,
//                               PT := T0S);
//                 END_IF;
//             END_IF;
//     END_CASE;
// {endregion}
// 
// {region "Shuttle Interlock"}
//     // VTD needs to be in Auto mode to perform a Shuttle interlock
//     CASE I_State OF
//         0:
//             IF VTD_Control.Mode = 3 AND VTD_Control.Shuttle_Interlock.Interlock_Request AND VTD_Control.Shuttle_Interlock.Shuttle_Interlock_Task_ID > 0 THEN
//                 I_State := 10;
//             END_IF;
//             
//         10: //Standby
//             
//             //Start by decoding all the IDs of the devices pertaining to the VTD in question on that level
//             "ID_Decode_F"(ID := VTD_Settings.ID,
//                           ID_Decoded := VTD_ID_Decoded);
//             "ID_Decode_F"(ID := "Settings_DB".LCnv_Sys[System_no].Cnv_Level[VTD_Control.Current_Level].Cnv1.ID,
//                           ID_Decoded := Cnv_ID_Decoded[1]);
//             "ID_Decode_F"(ID := "Settings_DB".LCnv_Sys[System_no].Cnv_Level[VTD_Control.Current_Level].Cnv2.ID,
//                           ID_Decoded := Cnv_ID_Decoded[2]);
//             
//             // Ensure the VTD is in a state that it can perform an interlock
//             IF VTD_Control.Docked AND NOT VTD_Control.Running AND (VTD_Control.Shuttle_Loaded = 0 OR VTD_Control.Shuttle_Loaded = 1) AND VTD_Control.Error = 0 THEN
//                 // Check to make sure the VTD and Shuttle are not both loaded
//                 IF VTD_Control.Pallet_Loaded = 1 THEN
//                     VTD_Control.Warning := 1; // Both the VTD and Shuttles are loaded, can't perform the interlock
//                 ELSE
//                     //Check that shuttle is on the correct floor, that the start location given and the shuttle actual position matches and the destination is the correct extractor barcode
//                     IF (*VTD_Control.Current_Level = "Shuttle_MQTT_DB".Shuttle_MQTT[VTD_Control.Shuttle_Interlock.Shuttle_ID].Message.Shuttle_Status.Floor
//                             AND*)VTD_Control.Shuttle_Interlock.Shuttle_Start_Location = "Shuttle_MQTT_DB".Shuttle_MQTT[VTD_Control.Shuttle_Interlock.Shuttle_ID].Message.Shuttle_Status.Position_ID
//                             (*AND "Shuttle_MQTT_DB".Shuttle_MQTT[VTD_Control.Shuttle_Interlock.Shuttle_ID].Message.Shuttle_Status.Destination_ID = "Settings_DB".ECnv_Settings.Barcode_ID*)THEN
//                         
//                         //Check in which Buffer conveyor the shuttle is located
//                         IF "Settings_DB".LCnv_Sys[System_no].Cnv_Level[VTD_Control.Current_Level].Cnv1.Barcode_ID =
//                             VTD_Control.Shuttle_Interlock.Shuttle_Start_Location THEN
//                             VTD_Control.Running := TRUE;
//                             I_State := 20;
//                         ELSIF "Settings_DB".LCnv_Sys[System_no].Cnv_Level[VTD_Control.Current_Level].Cnv2.Barcode_ID =
//                             VTD_Control.Shuttle_Interlock.Shuttle_Start_Location THEN
//                             VTD_Control.Running := TRUE;
//                             I_State := 25;
//                         ELSIF "Settings_DB".ECnv_Sys[System_no].Barcode_ID =
//                             VTD_Control.Shuttle_Interlock.Shuttle_Start_Location AND
//                             Control_GVL.VTD_Order_Table[System_no].Destination_Location = "Settings_DB".LCnv_Sys[System_no].Cnv_Level[VTD_Control.Current_Level].Cnv1.Barcode_ID THEN
//                             VTD_Control.Running := TRUE;
//                             I_State := 20;
//                         ELSIF "Settings_DB".ECnv_Sys[System_no].Barcode_ID =
//                             VTD_Control.Shuttle_Interlock.Shuttle_Start_Location AND
//                             Control_GVL.VTD_Order_Table[System_no].Destination_Location = "Settings_DB".LCnv_Sys[System_no].Cnv_Level[VTD_Control.Current_Level].Cnv2.Barcode_ID THEN
//                             VTD_Control.Running := TRUE;
//                             I_State := 25;
//                         ELSE
//                             VTD_Control.Warning := 2; // Shuttle interlock start location not buffer conveyor of VTD
//                         END_IF;
//                     ELSE
//                         VTD_Control.Warning := 3; // Cant interlock as shuttle and VTD level mismatch
//                     END_IF;
//                 END_IF;
//             ELSE
//                 VTD_Control.Warning := 4; // VTD not ready for interlock 
//             END_IF;
//             
//             
//         20: //Drop safety stops
//             IF Cnv_ID_Decoded[1].Level = VTD_Control.Current_Level THEN
//                 Control.LCnv_Sys[System_no].Cnv_Level[VTD_Control.Current_Level].Cnv1.Safety_Stop_Cnrl.Instruction.Retract := TRUE;
//                 I_State := 30;
//             ELSE
//                 VTD_Control.Error := TRUE; //24:16 Cannot find the correct safety pins to drop.
//                 Set_Bit_F(Bit_Number := 1,
//                             Bit_Value := 1,
//                             Variavel := VTD_Control.VTD_Errors.Error_Word_3);
//                 // I_State := 400;
//             END_IF;
//             
//         25: //Drop safety pins   
//             IF Cnv_ID_Decoded[2].Level = VTD_Control.Current_Level THEN
//                 Control.LCnv_Sys[System_no].Cnv_Level[VTD_Control.Current_Level].Cnv2.Safety_Stop_Cnrl.Instruction.Retract := TRUE;
//                 I_State := 35;
//             ELSE
//                 VTD_Control.Error := TRUE; //24:16 Cannot find the correct safety pins to drop.
//                 Set_Bit_F(Bit_Number := 1,
//                             Bit_Value := 1,
//                             Variavel := VTD_Control.VTD_Errors.Error_Word_3);
//                 // I_State := 400;
//             END_IF;
//             //////////////////////////////////////////////////////////////////////////////////////////////////////////////////////////////////////////////////////////////////    
//         30: //Confirm safety stops are down at the correct location
//             //Send ready to interlock
//             IF Control.LCnv_Sys[System_no].Cnv_Level[VTD_Control.Current_Level].Cnv1.Safety_Stop_Cnrl.LP_State = 0 THEN //RETRACTED
//                 Control.LCnv_Sys[System_no].Cnv_Level[VTD_Control.Current_Level].Cnv1.Safety_Stop_Cnrl.Instruction.Retract := FALSE;
//                 VTD_Control.Shuttle_Interlock.Ready_To_Interlock := TRUE;
//                 I_State := 40;
//             END_IF;
//             
//         35: //Confirm safety stops are down at the correct location
//             //Send ready to interlock
//             IF Control.LCnv_Sys[System_no].Cnv_Level[VTD_Control.Current_Level].Cnv2.Safety_Stop_Cnrl.LP_State = 0 THEN //RETRACTED
//                 Control.LCnv_Sys[System_no].Cnv_Level[VTD_Control.Current_Level].Cnv2.Safety_Stop_Cnrl.Instruction.Retract := FALSE;
//                 VTD_Control.Shuttle_Interlock.Ready_To_Interlock := TRUE;
//                 I_State := 45;
//             END_IF;
//             ////////////////////////////////////////////////////////////////////////////////////////////////////////////////////////////////////////////////////////////////////
//         40: //Wait for shuttle to move in or out VTD
//             IF Control_GVL.VTD_Order_Table[System_no].Destination_Location = "Settings_DB".ECnv_Sys[System_no].Barcode_ID THEN
//                 IF "Settings_DB".ECnv_Sys[System_no].Barcode_ID = "Shuttle_MQTT_DB".Shuttle_MQTT[VTD_Control.Shuttle_Interlock.Shuttle_ID].Message.Shuttle_Status.Position_ID
//                     AND "Shuttle_MQTT_DB".Shuttle_MQTT[VTD_Control.Shuttle_Interlock.Shuttle_ID].Message.Shuttle_Status.Operational_State = 'IDLE' THEN
//                     Control.LCnv_Sys[System_no].Cnv_Level[VTD_Control.Current_Level].Cnv1.Safety_Stop_Cnrl.Instruction.Extend := TRUE;
//                     I_State := 50;
//                 END_IF;
//             ELSIF Control.VTD_Order_Table[System_no].Destination_Location = "Settings_DB".LCnv_Sys[System_no].Cnv_Level[VTD_Control.Current_Level].Cnv1.Barcode_ID THEN
//                 IF "Settings_DB".LCnv_Sys[System_no].Cnv_Level[VTD_Control.Current_Level].Cnv1.Barcode_ID = "Shuttle_MQTT_DB".Shuttle_MQTT[VTD_Control.Shuttle_Interlock.Shuttle_ID].Message.Shuttle_Status.Position_ID
//                     AND "Shuttle_MQTT_DB".Shuttle_MQTT[VTD_Control.Shuttle_Interlock.Shuttle_ID].Message.Shuttle_Status.Operational_State = 'IDLE' THEN
//                     Control.LCnv_Sys[System_no].Cnv_Level[VTD_Control.Current_Level].Cnv1.Safety_Stop_Cnrl.Instruction.Extend := TRUE;
//                     I_State := 50;
//                 END_IF;
//             END_IF;
//             
//         45: //Wait for shuttle to move in or out VTD
//             IF Control_GVL.VTD_Order_Table[System_no].Destination_Location = "Settings_DB".ECnv_Sys[System_no].Barcode_ID THEN
//                 IF "Settings_DB".ECnv_Sys[System_no].Barcode_ID = "Shuttle_MQTT_DB".Shuttle_MQTT[VTD_Control.Shuttle_Interlock.Shuttle_ID].Message.Shuttle_Status.Position_ID
//                     AND "Shuttle_MQTT_DB".Shuttle_MQTT[VTD_Control.Shuttle_Interlock.Shuttle_ID].Message.Shuttle_Status.Operational_State = 'IDLE' THEN
//                     Control.LCnv_Sys[System_no].Cnv_Level[VTD_Control.Current_Level].Cnv2.Safety_Stop_Cnrl.Instruction.Extend := TRUE;
//                     I_State := 55;
//                 END_IF;
//             ELSIF Control.VTD_Order_Table[System_no].Destination_Location = "Settings_DB".LCnv_Sys[System_no].Cnv_Level[VTD_Control.Current_Level].Cnv2.Barcode_ID THEN
//                 IF "Settings_DB".LCnv_Sys[System_no].Cnv_Level[VTD_Control.Current_Level].Cnv2.Barcode_ID = "Shuttle_MQTT_DB".Shuttle_MQTT[VTD_Control.Shuttle_Interlock.Shuttle_ID].Message.Shuttle_Status.Position_ID
//                     AND "Shuttle_MQTT_DB".Shuttle_MQTT[VTD_Control.Shuttle_Interlock.Shuttle_ID].Message.Shuttle_Status.Operational_State = 'IDLE' THEN
//                     Control.LCnv_Sys[System_no].Cnv_Level[VTD_Control.Current_Level].Cnv2.Safety_Stop_Cnrl.Instruction.Extend := TRUE;
//                     I_State := 55;
//                 END_IF;
//             END_IF;
//             //////////////////////////////////////////////////////////////////////////////////////////////////////////////////////////////////////////////////////////////////////////  
//         50: //Check own sensors for shuttle/pallet state
//             IEC_Timer_0_Instance_1(IN := TRUE,
//                                     PT := T5S);
//             IF Control.LCnv_Sys[System_no].Cnv_Level[VTD_Control.Current_Level].Cnv1.Safety_Stop_Cnrl.LP_State = 1 //EXTENDED
//                 THEN
//                 Control.LCnv_Sys[System_no].Cnv_Level[VTD_Control.Current_Level].Cnv1.Safety_Stop_Cnrl.Instruction.Extend := FALSE;
//                 VTD_Control.Shuttle_Interlock.Interlock_Complete := TRUE;
//                 I_State := 60;
//             ELSIF IEC_Timer_0_Instance_1.Q THEN
//                 VTD_Control.Error := TRUE; //24:17 Error occured during interlock final check
//                 Set_Bit_F(Bit_Number := 2,
//                             Bit_Value := 1,
//                             Variavel := VTD_Control.VTD_Errors.Error_Word_3);
//                 I_State := 400;
//             END_IF;
//             
//         55: //Check own sensors for shuttle/pallet state
//             IEC_Timer_0_Instance_1(IN := TRUE,
//                                     PT := T5S);
//             IF Control.LCnv_Sys[System_no].Cnv_Level[VTD_Control.Current_Level].Cnv2.Safety_Stop_Cnrl.LP_State = 1 //EXTENDED
//                 THEN
//                 Control.LCnv_Sys[System_no].Cnv_Level[VTD_Control.Current_Level].Cnv2.Safety_Stop_Cnrl.Instruction.Extend := FALSE;
//                 VTD_Control.Shuttle_Interlock.Interlock_Complete := TRUE;
//                 I_State := 60;
//             ELSIF IEC_Timer_0_Instance_1.Q THEN
//                 VTD_Control.Error := TRUE; //24:17 Error occured during interlock final check
//                 Set_Bit_F(Bit_Number := 2,
//                             Bit_Value := 1,
//                             Variavel := VTD_Control.VTD_Errors.Error_Word_3);
//                 I_State := 400;
//             END_IF;
//             
//         60://Clear Vars
//             IEC_Timer_0_Instance_1(IN := FALSE,
//                                     PT := T0s);
//             IEC_Timer_0_Instance_2(IN := FALSE,
//                                     PT := T0s);
//             IF VTD_Control.Shuttle_Interlock.Interlock_Complete_Ack THEN
//                 VTD_Control.Shuttle_Interlock.Ready_To_Interlock := FALSE;
//                 VTD_Control.Shuttle_Interlock.Interlock_Complete := FALSE;
//                 VTD_Control.Running := FALSE;
//                 I_State := 0;
//             END_IF;
//             
//         400://ERROR MODE
//             IEC_Timer_0_Instance_1(IN := FALSE,
//                                     PT := T#0S);
//             IEC_Timer_0_Instance_2(IN := FALSE,
//                                     PT := T#0S);
//             Interlock_Timer(IN := FALSE,
//                              PT := T#0S);
//             VTD_Control.Running := FALSE;
//             VTD_Control.Shuttle_Interlock.Interlock_Complete := FALSE;
//             VTD_Control.Shuttle_Interlock.Ready_To_Interlock := FALSE;
//             Control.LCnv_Sys[System_no].Cnv_Level[VTD_Control.Current_Level].Cnv1.Safety_Stop_Cnrl.Instruction.Extend := FALSE;
//             Control.LCnv_Sys[System_no].Cnv_Level[VTD_Control.Current_Level].Cnv2.Safety_Stop_Cnrl.Instruction.Extend := FALSE;
//             Control.LCnv_Sys[System_no].Cnv_Level[VTD_Control.Current_Level].Cnv1.Safety_Stop_Cnrl.Instruction.Retract := FALSE;
//             Control.LCnv_Sys[System_no].Cnv_Level[VTD_Control.Current_Level].Cnv2.Safety_Stop_Cnrl.Instruction.Retract := FALSE;
//             IF VTD_Control.Instruction.Reset THEN
//                 VTD_Control.VTD_Errors.Error_Word_3 := 0;
//                 I_State := 0;
//             END_IF;
//     END_CASE;
//     Interlock_Timer(IN := I_State >= 40 AND I_State <= 50,
//                      PT := UINT_TO_TIME("Settings_DB".System.Shuttle_Interlock_Timeout) * 1000);
//     
// {endregion}
// 
// 
// // IF System_no <> 3 THEN
// {region "Cyclic Error Checks"}
//     IF NOT Safety_OK THEN //SAFETY
//         Set_Bit_F(Bit_Number := 0,
//                   Variavel := VTD_Control.VTD_Errors.Error_Word_1);
//     END_IF;
//     
//     IF VTD_Control.Instruction.Stop THEN //HMI STOP
//         Set_Bit_F(Bit_Number := 1,
//                     Variavel := VTD_Control.VTD_Errors.Error_Word_1);
//     END_IF;
//     
//     IF NOT VTD_Control.Inputs.Upper_Overtravel AND NOT Bypass.Upper_limit THEN //UPPER OVERTRAVEL
//         Set_Bit_F(Bit_Number := 2,
//                     Variavel := VTD_Control.VTD_Errors.Error_Word_1);
//     END_IF;
//     
//     IF NOT VTD_Control.Inputs.Lower_Overtravel AND NOT Bypass.Lower_limit THEN //LOWER OVERTRAVEL
//         Set_Bit_F(Bit_Number := 3,
//                     Variavel := VTD_Control.VTD_Errors.Error_Word_1);
//     END_IF;
//     
//     //CHAIN SLACK
//     IF Chain_Slack_1 AND NOT Bypass.Chain_Slack_1 THEN
//         Set_Bit_F(Bit_Number := 0,
//                     Variavel := VTD_Control.VTD_Errors.Error_Word_5);
//     END_IF;
//     
//     IF Chain_Slack_2 AND NOT Bypass.Chain_Slack_2 THEN
//         Set_Bit_F(Bit_Number := 1,
//                     Variavel := VTD_Control.VTD_Errors.Error_Word_5);
//     END_IF;
//     
//     IF Chain_Slack_3 AND NOT Bypass.Chain_Slack_3 THEN
//         Set_Bit_F(Bit_Number := 2,
//                     Variavel := VTD_Control.VTD_Errors.Error_Word_5);
//     END_IF;
//     
//     IF Chain_Slack_4 AND NOT Bypass.Chain_Slack_4 THEN
//         Set_Bit_F(Bit_Number := 3,
//                     Variavel := VTD_Control.VTD_Errors.Error_Word_5);
//     END_IF;
//     
//     //VFD ERROR
//     IF fbSewDrive.q_bError THEN // SEW: drive fault or communication error
//         Set_Bit_F(Bit_Number := 7,
//                     Variavel := VTD_Control.VTD_Errors.Error_Word_4);
//     END_IF;
//     
//     //HIGH LIMITS
//     IF VTD_Control.LinearEnc > VTD_Settings.VTD_Max_Heigh AND NOT LE_Bypass_HMI AND NOT "VTD_HMI".LE_Bypass[System_no] THEN //21:5
//         Set_Bit_F(Bit_Number := 4,
//                     Variavel := VTD_Control.VTD_Errors.Error_Word_1);
//     END_IF;
//     
//     IF VTD_Control.LinearEnc < VTD_Settings.VTD_Min_Height AND NOT LE_Bypass_HMI AND NOT "VTD_HMI".LE_Bypass[System_no] THEN //21:5
//         Set_Bit_F(Bit_Number := 5,
//                     Variavel := VTD_Control.VTD_Errors.Error_Word_1);
//     END_IF;
//     
//     //AUTOMATIC MODE NOT DOCKED
//     R_AutomatcMode(CLK := VTD_Control.Mode = 3);
//     IF NOT VTD_Control.Docked AND R_AutomatcMode.Q THEN //22:1
//         Set_Bit_F(Bit_Number := 8,
//                     Variavel := VTD_Control.VTD_Errors.Error_Word_1);
//     END_IF;
//     
//     IF NOT Level_Detect AND R_AutomatcMode.Q THEN //22:2
//         Set_Bit_F(Bit_Number := 9,
//                     Variavel := VTD_Control.VTD_Errors.Error_Word_1);
//     END_IF;
//     
//     //TRYING RETRACT WHILE DOCKED
//     IF VTD_Control.Docked AND (DP1_Retract OR DP2_Retract) THEN //22:5
//         Set_Bit_F(Bit_Number := 12,
//                     Variavel := VTD_Control.VTD_Errors.Error_Word_1);
//     END_IF;
//     
//     //LE ERROR
//     T_LE_Error.TON(IN := VTD_Control.Inputs.LE_Status.%X0 OR VTD_Control.Inputs.LE_Status.%X1 OR
//                     VTD_Control.LinearEnc < VTD_Settings.VTD_Min_Height OR
//                     VTD_Control.LinearEnc > VTD_Settings.VTD_Max_Heigh,
//                     PT := t500ms);
//     IF NOT LE_Bypass_HMI AND NOT "VTD_HMI".LE_Bypass[System_no] AND T_LE_Error.Q THEN
//         Set_Bit_F(Bit_Number := 4,
//                     Variavel := VTD_Control.VTD_Errors.Error_Word_3);
//         T_LE_Error.TON(IN := FALSE,
//                         PT := T0s);
//     END_IF;
//     
//     
//     
//     //ABSOLUTE ENCODER
//     IF VTD_Control.AE_Error > 0 THEN
//         Set_Bit_F(Bit_Number := 5,
//                     Variavel := VTD_Control.VTD_Errors.Error_Word_3);
//         VTD_Control.Outputs.AE_Control_Word_1.7 := VTD_Control.Instruction.Reset OR Reset_All OR HMI_Reset;
//     ELSE
//         VTD_Control.Outputs.AE_Control_Word_1.7 := FALSE;
//     END_IF;
//     
//     IEC_Timer_0_Instance(IN := VTD_Control.LinearEnc <= (VTD_Settings.Teach_Values.Levels_LE[LevelBelowExtractor] + 1) AND VTD_Control.Instruction.Manual_Down,
//                           PT := T#300MS);
//     
//     //Errors while running
//     IF VTD_Control.Running THEN
//         IF LevelBelowExtractor < 7 THEN
//             IF NOT (VTD_Control.LP_State = 2) AND // NOT 'Retracted'
//                 (VTD_Control.LinearEnc > (VTD_Settings.Teach_Values.Levels_LE[LevelBelowExtractor] + VTD_Settings.Slowdown_Count_LE) AND
//                 VTD_Control.LinearEnc < (VTD_Settings.Teach_Values.Levels_LE[LevelBelowExtractor + 1] - VTD_Settings.Creep_Count_LE) AND
//                 VTD_Control.Instruction.Manual_Up)
//                 OR
//                 IEC_Timer_0_Instance.Q
//             THEN //22:4
//                 IF NOT Bypass_LP THEN
//                     IF System_no <> 5 THEN
//                         Set_Bit_F(Bit_Number := 11,
//                                     Variavel := VTD_Control.VTD_Errors.Error_Word_1);
//                     END_IF;
//                 END_IF;
//             END_IF;
//         ELSIF LevelBelowExtractor = 8 THEN
//             IF NOT (VTD_Control.LP_State = 2) AND // NOT 'Retracted'
//                 (VTD_Control.LinearEnc > (VTD_Settings.Teach_Values.Levels_LE[LevelBelowExtractor] + VTD_Settings.Slowdown_Count_LE) AND
//                 VTD_Control.Instruction.Manual_Up)
//                 OR
//                 IEC_Timer_0_Instance.Q
//             THEN //22:4
//                 IF NOT Bypass_LP THEN
//                     IF System_no <> 5 THEN
//                         Set_Bit_F(Bit_Number := 11,
//                                     Variavel := VTD_Control.VTD_Errors.Error_Word_1);
//                     END_IF;
//                 END_IF;
//             END_IF;
//         END_IF;
//         
//         IF fbSewDrive.q_bError THEN //VFD ERROR (SEW: drive fault or communication error)
//             Set_Bit_F(Bit_Number := 0,
//                         Variavel := VTD_Control.VTD_Errors.Error_Word_4);
//         ELSIF VTD_Control.LinearEnc_Error > 0 THEN //LE ERROR
//             Set_Bit_F(Bit_Number := 1,
//                         Variavel := VTD_Control.VTD_Errors.Error_Word_4);
//         ELSIF VTD_Control.AE_Error > 0 THEN //AE ERROR
//             Set_Bit_F(Bit_Number := 2,
//                         Variavel := VTD_Control.VTD_Errors.Error_Word_4);
//             
//         ELSIF (DP1_Extended AND DP1_Retracted) OR (DP2_Extended AND DP2_Retracted) THEN // 25:4
//             IF System_no <> 5 THEN
//                 Set_Bit_F(Bit_Number := 3,
//                             Variavel := VTD_Control.VTD_Errors.Error_Word_4);
//             ELSE
//                 ;
//             END_IF;
//         ELSIF Lower_Limit AND NOT Upper_limit AND NOT Bypass.Overtravel_Lower_limit THEN // 25:5
//             Set_Bit_F(Bit_Number := 4,
//                         Variavel := VTD_Control.VTD_Errors.Error_Word_4);
//         ELSIF NOT Lower_Limit AND Upper_limit AND NOT Bypass.Overtravel_Upper_limit THEN // 25:6
//             Set_Bit_F(Bit_Number := 5,
//                         Variavel := VTD_Control.VTD_Errors.Error_Word_4);
//         ELSIF Lower_Limit AND Upper_limit THEN // 25:7
//             Set_Bit_F(Bit_Number := 6,
//                         Variavel := VTD_Control.VTD_Errors.Error_Word_4);
//         END_IF;
//     END_IF;
//     
//     //Check if overtravel limit switches has been hit
//     IF Upper_limit AND VTD_Control.Instruction.Manual_Up
//     THEN //24:6 Top overtravel limit reached.
//         Set_Bit_F(Bit_Number := 7,
//                     Variavel := VTD_Control.VTD_Errors.Error_Word_2);
//         IF VTD_Control.Mode = 2 OR VTD_Control.Mode = 3 THEN
//             State := 400;
//         ELSE
//             State := 0;
//         END_IF;
//     ELSIF Lower_Limit AND VTD_Control.Instruction.Manual_Down
//     THEN //24:7 Bottom overtravel limit reached.
//         Set_Bit_F(Bit_Number := 8,
//                     Variavel := VTD_Control.VTD_Errors.Error_Word_2);
//         IF VTD_Control.Mode = 2 OR VTD_Control.Mode = 3 THEN
//             State := 400;
//         ELSE
//             State := 0;
//         END_IF;
//     END_IF;
//     
//     //Need to monitor both encoders
//     IF ABS(VTD_Control.Encoder_Delta) > VTD_Settings.Encoder_Delta_Warning THEN
//         VTD_Control.Warning := 2;
//     END_IF;
//     
//     T_Encoders_Difference(IN := ABS(VTD_Control.Encoder_Delta) > VTD_Settings.Encoder_Delta_Error,
//                            PT := T#500MS);
//     
//     IF T_Encoders_Difference.Q AND NOT LE_Bypass_HMI AND NOT "VTD_HMI".LE_Bypass[System_no] THEN
//         //Send error message that encoder error is to large
//         Set_Bit_F(Bit_Number := 2,
//                     Variavel := VTD_Control.VTD_Errors.Error_Word_2);
//     END_IF;
//     
//     // Level detect timer 
//     IF LD_Timer.Q OR LD_Timer_1.Q THEN
//         LD_Timer(IN := FALSE,
//                   PT := T#0S);
//         LD_Timer_1(IN := FALSE,
//                     PT := T#0S);
//             Set_Bit_F(Bit_Number := 11,
//                         Variavel := VTD_Control.VTD_Errors.Error_Word_4);
//     END_IF;
//     
//     //Locking pin timer
//     IF DP_Timer.Q AND (DP1_Retract OR DP1_Extend) THEN //24:2 Locking pins took to long to extend
//         Set_Bit_F(Bit_Number := 3,
//                     Variavel := VTD_Control.VTD_Errors.Error_Word_2);
//     ELSIF DP_Timer.Q AND (DP2_Retract AND DP2_Extend) THEN //24:3 Locking pins took to long to retract
//         Set_Bit_F(Bit_Number := 4,
//                     Variavel := VTD_Control.VTD_Errors.Error_Word_2);
//     END_IF;
//     
//     IF Interlock_Timer.Q THEN //Interlock process timed out
//         Set_Bit_F(Bit_Number := 3,
//                     Variavel := VTD_Control.VTD_Errors.Error_Word_3);
//         I_State := 400;
//     END_IF;
//     
//     //MOVIVENT VTD UNEXPECTED
//     //Take the position old
//     R_Position_OLD(CLK:= NOT VTD_Control.Motor_UP AND NOT VTD_Control.Motor_Down AND MainSetpoint1 = 0);
//     
//     IF R_Position_OLD.Q THEN
//         Position_OLD := VTD_Control.LinearEnc;
//     ELSIF NOT R_Position_OLD.CLK THEN
//         Position_OLD := 0;
//     END_IF;
//     
//     //VTD STILL MOVING
//     IF ABS(VTD_Control.LinearEnc - Position_OLD) > Tol_VTD_Still_Moving THEN
//         Set_Bit_F(Bit_Number := 6,
//                     Variavel := VTD_Control.VTD_Errors.Error_Word_3);
//     END_IF;
//     
//     // Watchdog bit
//     // IF Watchdog.Q THEN
//     //     VTD_Control.Running := FALSE;
//     //     IF VTD_Control.Mode = 4 THEN //24:9 Teach timed out
//     //         Set_Bit_F(Bit_Number := 10,
//     //                     Bit_Value := 1,
//     //                     Variavel := VTD_Control.VTD_Errors.Error_Word_2);
//     //     ELSIF VTD_Control.Mode = 3 THEN //24:9 Auto timed out
//     //         Set_Bit_F(Bit_Number := 10,
//     //                     Bit_Value := 1,
//     //                     Variavel := VTD_Control.VTD_Errors.Error_Word_2);
//     //     ELSIF VTD_Control.Mode = 2 THEN //24:9 Semi auto timed out
//     //         Set_Bit_F(Bit_Number := 10,
//     //                     Bit_Value := 1,
//     //                     Variavel := VTD_Control.VTD_Errors.Error_Word_2);
//     //     END_IF;
//     // END_IF;
//     
//     IF ((System_no = 1 AND "Errors_Profinet_1".%X8) OR
//         (System_no = 2 AND "Errors_Profinet_3".%X7) OR
//         (System_no = 3 AND "Errors_Profinet_5".%X4) OR
//         (System_no = 4 AND "Errors_Profinet_7".%X1) OR
//         (System_no = 5 AND "Errors_Profinet_8".%X6)) AND VTD_Control.Mode = 3
//     THEN //Interface Profinet error
//         Set_Bit_F(Bit_Number := 3,
//                     Variavel := VTD_Control.VTD_Errors.Error_Word_3);
//     END_IF;
//     
//     // go to error state
//     IF VTD_Control.VTD_Errors.Error_Word_1 <> 0 OR
//         VTD_Control.VTD_Errors.Error_Word_2 <> 0 OR
//         VTD_Control.VTD_Errors.Error_Word_3 <> 0 OR
//         VTD_Control.VTD_Errors.Error_Word_4 <> 0 OR
//         VTD_Control.VTD_Errors.Error_Word_5 <> 0 THEN
//         VTD_Control.Error := TRUE;
//         State := 400;
//     END_IF;
// {endregion}
// // END_IF;
// 
{region "VFD - SEW MOVIPRO, MOVIKIT Positioning Drive, speed mode (200)"}
    // Adapted from the former G120/SinaSpeed region. The state machine above still
    // commands the motor exactly as before:
    //   VTD_Control.Motor_UP / Motor_Down = direction
    //   VTD_Control.Motor_Speed           = speed in % (0..120), 100 % = VTD_Settings.SEW_Speed_At_100pct
    // This region converts those commands to MOVIKIT speed mode (200), SEW manual 33959862, 8.1.4.
    // ASSUMPTION (verify on the first test): a positive speed setpoint moves the VTD up.
    // If not, correct the direction of rotation in MOVISUITE, not here.

    //SETPOINT (signed, user units)
    IF VTD_Control.Motor_UP AND NOT VTD_Control.Motor_Down THEN
        rSpeedSetpoint := UINT_TO_REAL(MIN(VTD_Control.Motor_Speed, 120))
                          * INT_TO_REAL(VTD_Settings.SEW_Speed_At_100pct) / 100.0;
    ELSIF VTD_Control.Motor_Down AND NOT VTD_Control.Motor_UP THEN
        rSpeedSetpoint := -1.0 * UINT_TO_REAL(MIN(VTD_Control.Motor_Speed, 120))
                          * INT_TO_REAL(VTD_Settings.SEW_Speed_At_100pct) / 100.0;
    ELSE
        rSpeedSetpoint := 0.0;
    END_IF
    MainSetpoint := REAL_TO_INT(LIMIT(-32767.0, rSpeedSetpoint, 32767.0));

    T_Setpoint_Delay(IN := MainSetpoint <> 0,
                     PT := T#0MS);

    IF T_Setpoint_Delay.Q THEN
        MainSetpoint1 := MainSetpoint;
    ELSE
        MainSetpoint1 := 0;
    END_IF

    //Acceleration: same load/weight ranges as before, as a factor in %
    diPalletWeight := 0;
    IF System_no >= 1 AND System_no <= 2 THEN // Control.VTD_Order_Table is ARRAY[1..2]
        diPalletWeight := INT_TO_DINT(Control.VTD_Order_Table.Pallet_Weight);
    END_IF

    IF VTD_Control.Pallet_Loaded = 0 AND VTD_Control.Shuttle_Loaded = 0 THEN
        rAccelerationFactor_pct := 60.0;
    ELSIF diPalletWeight > 0 AND diPalletWeight <= UINT_TO_DINT(VTD_Settings.Weight_Range_1) THEN
        rAccelerationFactor_pct := UINT_TO_REAL(VTD_Settings.Acc_Range_1);
    ELSIF diPalletWeight > UINT_TO_DINT(VTD_Settings.Weight_Range_1)
        AND diPalletWeight <= UINT_TO_DINT(VTD_Settings.Weight_Range_2) THEN
        rAccelerationFactor_pct := UINT_TO_REAL(VTD_Settings.Acc_Range_2);
    ELSIF diPalletWeight > UINT_TO_DINT(VTD_Settings.Weight_Range_2)
        AND diPalletWeight <= UINT_TO_DINT(VTD_Settings.Weight_Range_3) THEN
        rAccelerationFactor_pct := UINT_TO_REAL(VTD_Settings.Acc_Range_3);
    ELSE
        rAccelerationFactor_pct := 100.0;
    END_IF

    uiDriveRamp := REAL_TO_UINT(LIMIT(0.0,
                                      rAccelerationFactor_pct * UINT_TO_REAL(VTD_Settings.SEW_Ramp_At_100pct) / 100.0,
                                      65535.0));

    //ENABLE / START
    bDriveMoveRequest := (VTD_Control.Motor_UP XOR VTD_Control.Motor_Down) AND MainSetpoint1 <> 0;

    // Keep the enable until the motor has stopped, so a normal stop (start = 0)
    // decelerates with the PO 4 ramp before the brake is applied.
    // Safety_OK or a VTD error removes the enable immediately (FCB 14 emergency stop ramp).
    bDriveEnable := Safety_OK AND NOT VTD_Control.Error
                    AND (bDriveMoveRequest OR VTD_Control.Motor.stStatus.bMotorTurning);

    bDriveFaultReset := VTD_Control.Instruction.Reset OR System_Control.Reset_All OR HMI_Reset;

    fbSewDrive(i_stProcessInput := VTD_Control.Motor.stProcessInput,
               i_bEnable := bDriveEnable,
               i_bStart := bDriveMoveRequest AND bDriveEnable,
               i_bJogPositive := FALSE,
               i_bJogNegative := FALSE,
               i_bFaultReset := bDriveFaultReset,
               i_eMode := E_SEW_MovikitMode.Speed,
               i_iSpeedSetpoint := MainSetpoint1,
               i_uiAcceleration := uiDriveRamp,
               i_uiDeceleration := uiDriveRamp,
               i_diTargetPosition := 0);

    VTD_Control.Motor.aProcessOutput := fbSewDrive.q_aProcessOutput;
    VTD_Control.Motor.stStatus := fbSewDrive.q_stStatus;

    //VFD error code: 16#FFFF = communication, otherwise PI 3 (fault * 256 + subfault)
    IF NOT fbSewDrive.q_stStatus.bCommunicationOk THEN
        VTD_Control.VFD_Error := 16#FFFF;
    ELSIF fbSewDrive.q_stStatus.bError THEN
        VTD_Control.VFD_Error := VTD_Control.Motor.stProcessInput.aWord[3];
    ELSE
        VTD_Control.VFD_Error := 0;
    END_IF

    // TODO: VTD_Control.LinearEnc [mm] from fbSewDrive.q_stStatus.diActualPosition (DL50 via PI 7/8)
    //       once the MOVISUITE user units of the position are confirmed.
{endregion}
// 
// HMI_Reset := (("Screen_DB_1".Reset_All[1] OR "VTD_HMI".Reset[1]) AND
// ("HMI_Box_Connected_1" = 11 AND "KEY REMOTE/LOCAL L1 - CH1(1)") OR
// ("HMI_Box_Connected_1" = 12 AND "KEY REMOTE/LOCAL L2 - CH1(1)") OR
// ("HMI_Box_Connected_1" = 13 AND "KEY REMOTE/LOCAL L3 - CH1(1)") OR
// ("HMI_Box_Connected_1" = 14 AND "KEY REMOTE/LOCAL L4 - CH1(1)") OR
// ("HMI_Box_Connected_1" = 15 AND "KEY REMOTE/LOCAL L5 - CH1(1)") OR
// ("HMI_Box_Connected_1" = 16 AND "KEY REMOTE/LOCAL L6 - CH1(1)") OR
// ("HMI_Box_Connected_1" = 21 AND "KEY REMOTE/LOCAL L1 - CH1(2)") OR
// ("HMI_Box_Connected_1" = 22 AND "KEY REMOTE/LOCAL L2 - CH1(2)") OR
// ("HMI_Box_Connected_1" = 23 AND "KEY REMOTE/LOCAL L3 - CH1(2)") OR
// ("HMI_Box_Connected_1" = 24 AND "KEY REMOTE/LOCAL L4 - CH1(2)") OR
// ("HMI_Box_Connected_1" = 25 AND "KEY REMOTE/LOCAL L5 - CH1(2)") OR
// ("HMI_Box_Connected_1" = 26 AND "KEY REMOTE/LOCAL L6 - CH1(2)"))
// OR
// (("Screen_DB_1".Reset_All[2] OR "VTD_HMI".Reset[2]) AND
// ("HMI_Box_Connected_2" = 11 AND "KEY REMOTE/LOCAL L1 - CH1(1)") OR
// ("HMI_Box_Connected_2" = 12 AND "KEY REMOTE/LOCAL L2 - CH1(1)") OR
// ("HMI_Box_Connected_2" = 13 AND "KEY REMOTE/LOCAL L3 - CH1(1)") OR
// ("HMI_Box_Connected_2" = 14 AND "KEY REMOTE/LOCAL L4 - CH1(1)") OR
// ("HMI_Box_Connected_2" = 15 AND "KEY REMOTE/LOCAL L5 - CH1(1)") OR
// ("HMI_Box_Connected_2" = 16 AND "KEY REMOTE/LOCAL L6 - CH1(1)") OR
// ("HMI_Box_Connected_2" = 21 AND "KEY REMOTE/LOCAL L1 - CH1(2)") OR
// ("HMI_Box_Connected_2" = 22 AND "KEY REMOTE/LOCAL L2 - CH1(2)") OR
// ("HMI_Box_Connected_2" = 23 AND "KEY REMOTE/LOCAL L3 - CH1(2)") OR
// ("HMI_Box_Connected_2" = 24 AND "KEY REMOTE/LOCAL L4 - CH1(2)") OR
// ("HMI_Box_Connected_2" = 25 AND "KEY REMOTE/LOCAL L5 - CH1(2)") OR
// ("HMI_Box_Connected_2" = 26 AND "KEY REMOTE/LOCAL L6 - CH1(2)"));
// 
// //Assign local vars to outputs
// VTD_Control.Outputs.LP1_Retract := DP1_Retract;
// VTD_Control.Outputs.LP1_Extend := DP1_Extend;
// VTD_Control.Outputs.LP2_Retract := DP2_Retract;
// VTD_Control.Outputs.LP2_Extend := DP2_Extend;

END_FUNCTION_BLOCK

// ---- GlobalTextList.TcGTLO
TEXTLIST GlobalTextList
  2214 = '   %s  |  ACCESS GATES'
  2222 = '   %s  |  ALARMS'
  2205 = '   %s  |  CAROUSEL'
  2181 = '   %s  |  CONVEYORS'
  2072 = '   %s  |  MAIN'
  2226 = '   %s  |  ORDER TABLE'
  2230 = '   %s  |  SHUTTLES'
  2123 = '   %s  |  VTD'
  2001 = '   VTD MOVIPRO - Manual Test (TEST ONLY)'
  2199 = '%.1f %%'
  2209 = '%.1f deg'
  2151 = '%.1f mm'
  2147 = '%.1f mm/s'
  2149 = '%.2f A'
  1019 = '%04X'
  2022 = '%08X'
  457 = '%d'
  2031 = '%d %%'
  1082 = '%s'
  2066 = '%t[mm:ss]'
  2073 = '%t[yyyy-MM-dd HH:mm:ss]'
  661 = '%u'
  2057 = '(not an emergency stop)'
  1034 = '(PI 7 + PI 8)'
  1038 = '0'
  1087 = '0 - Ready'
  2069 = '0 = not configured: no motion accepted.'
  1039 = '1'
  2023 = '1 - Operating mode (changes only at standstill)'
  1088 = '1 - STO inactive'
  1048 = '10'
  2033 = '10 %'
  1097 = '10 - Drive train 2 active'
  2036 = '100 %'
  2038 = '100 % ='
  1049 = '11'
  1098 = '11 - Speed reached'
  1050 = '12'
  1099 = '12 - SW limit switches inactive'
  1051 = '13'
  1100 = '13 - Reserved'
  1052 = '14'
  1101 = '14 - Standby active'
  1053 = '15'
  1102 = '15 - Handshake Out'
  1040 = '2'
  1089 = '2 - Output stage enabled'
  2030 = '2 - Speed (% of the max test speed)'
  2034 = '25 %'
  1041 = '3'
  1090 = '3 - Brake released'
  2040 = '3 - Motion'
  1042 = '4'
  1091 = '4 - Motor turning'
  1043 = '5'
  2032 = '5 %'
  1092 = '5 - Referenced'
  2035 = '50 %'
  1044 = '6'
  1093 = '6 - New relative position applied'
  1045 = '7'
  1094 = '7 - In position'
  1046 = '8'
  1095 = '8 - Error'
  1047 = '9'
  1096 = '9 - Warning'
  2002 = '<< Process data'
  2071 = '>> Manual test'
  2131 = 'A'
  2138 = 'Abs. encoder'
  2063 = 'Acceleration'
  2118 = 'ACCESS GATES'
  2218 = 'Access granted'
  2217 = 'Access requested'
  2079 = 'Active alarms'
  1029 = 'Actual application mode'
  1081 = 'Actual mode'
  2018 = 'Actual mode (PI 6)'
  1002 = 'Actual position (DL50 via PI 7 high + PI 8 low)'
  1031 = 'Actual position - high word'
  1033 = 'Actual position - low word'
  1021 = 'Actual speed'
  2014 = 'Actual values (user units)'
  2142 = 'AE err.'
  2225 = 'Alarm source not defined yet (TwinCAT EventLogger or own alarm table).'
  2223 = 'Alarms'
  2080 = 'ALARMS'
  2224 = 'ALARMS - screen in preparation'
  1054 = 'Allow control word (PO 1)'
  2060 = 'and clears the software stop'
  2208 = 'Angle'
  2075 = 'Auto mode'
  2202 = 'BACKWARD'
  2194 = 'Backward sensor'
  2140 = 'Barcode'
  2008 = 'Brake released'
  2108 = 'Buffer L1'
  2107 = 'Buffer L2'
  2106 = 'Buffer L3'
  2105 = 'Buffer L4'
  2104 = 'Buffer L5'
  2103 = 'Buffer L6'
  2117 = 'CAROUSEL'
  2091 = 'Chain'
  2070 = 'Check the user units in MOVISUITE first.'
  2143 = 'Code err.'
  193 = 'Communication'
  1008 = 'Communication OK'
  1062 = 'Control word'
  2116 = 'CONVEYORS'
  2148 = 'Current'
  2134 = 'Current level'
  2132 = 'Data'
  2064 = 'Deceleration'
  1016 = 'Decoded'
  2183 = 'Device'
  2182 = 'Devices'
  1027 = 'Digital inputs'
  1079 = 'Digital inputs (PI 5)'
  1070 = 'Digital outputs'
  2196 = 'Direction'
  2128 = 'Docked'
  2137 = 'Docking pins'
  2215 = 'Door closed'
  2216 = 'Door locked'
  2161 = 'DP1 ext.'
  2163 = 'DP1 retr.'
  2162 = 'DP2 ext.'
  2164 = 'DP2 retr.'
  2144 = 'Drive'
  2054 = 'Drive commands'
  2012 = 'Drive error'
  2004 = 'Drive status (PI 1)'
  1055 = 'Elapsed %t[mm:ss]'
  2184 = 'En'
  2055 = 'ENABLE'
  2126 = 'Enabled'
  2139 = 'Encoder delta'
  2185 = 'Err'
  2078 = 'Error'
  2021 = 'Error ID (hex)'
  1010 = 'EtherCAT state'
  1012 = 'EtherCAT state 8 = OP. The counter must keep rising while the drive is powered.'
  2109 = 'Extractor'
  2020 = 'Fault / subfault'
  2203 = 'FORWARD'
  2193 = 'Forward sensor'
  2201 = 'From ID'
  2094 = 'Gate 1'
  2095 = 'Gate 2'
  2043 = 'hold to run'
  2011 = 'In position'
  2042 = 'JOG +'
  2041 = 'JOG -'
  2204 = 'Jog buttons: hold to run, manual mode only.'
  2065 = 'Jog max time'
  2025 = 'JOG position - 100'
  2024 = 'JOG speed - 101'
  2052 = 'JOG, RUN and START need ENABLE. Reversing in mode 200: press STOP first.'
  2141 = 'LE err.'
  2150 = 'LE position'
  2152 = 'LE speed'
  2180 = 'Level'
  2178 = 'Level 1'
  2177 = 'Level 2'
  2176 = 'Level 3'
  2175 = 'Level 4'
  2174 = 'Level 5'
  2173 = 'Level 6'
  2172 = 'Level 7'
  2171 = 'Level 8'
  2135 = 'Level below'
  2155 = 'Level det. 1'
  2156 = 'Level det. 2'
  2207 = 'Lift down'
  2210 = 'LIFT DOWN'
  2206 = 'Lift up'
  2211 = 'LIFT UP'
  2179 = 'Lower limit'
  2129 = 'M'
  2124 = 'MAIN'
  2076 = 'Manual mode'
  2121 = 'MANUAL TEST'
  2062 = 'Max speed (100 %)'
  1058 = 'Meaning'
  1014 = 'Meaning (MOVISUITE)'
  2235 = 'MENU'
  2046 = 'mode 200'
  2053 = 'Mode buttons are locked while the axis moves or a motion command is active.'
  2019 = 'Mode sent to the drive (PO 6)'
  2153 = 'Motor ready'
  2009 = 'Motor turning'
  891 = 'Open dialog'
  2229 = 'Order structure (OrderTable_DUT / WMS) to be confirmed.'
  2119 = 'ORDER TABLE'
  2227 = 'Order Table'
  2228 = 'ORDER TABLE - screen in preparation'
  2169 = 'OT limit'
  2007 = 'Output stage enabled'
  2186 = 'Pal'
  2112 = 'Pallet present'
  2133 = 'Pallet type'
  1017 = 'PI 1'
  1020 = 'PI 2'
  1022 = 'PI 3'
  1085 = 'PI 3: high byte = fault, low byte = subfault (active FCB if no fault).'
  1024 = 'PI 4'
  1026 = 'PI 5'
  1028 = 'PI 6'
  1030 = 'PI 7'
  1032 = 'PI 8'
  1011 = 'PI change counter'
  1061 = 'PO 1'
  1063 = 'PO 2'
  2037 = 'PO 2 sent'
  1065 = 'PO 3'
  1067 = 'PO 4'
  1069 = 'PO 5'
  1071 = 'PO 6'
  1073 = 'PO 7'
  1075 = 'PO 8'
  2084 = 'PopUp 1'
  2085 = 'PopUp 2'
  2028 = 'POS ABSOLUTE - 400'
  2029 = 'POS RELATIVE - 401'
  2015 = 'Position'
  2122 = 'PROCESS DATA'
  1077 = 'Process inputs (drive -> PLC)'
  1015 = 'Raw (hex)'
  2068 = 'Raw PD write active (process data screen)'
  1036 = 'Raw user units'
  1007 = 'Raw write: PO 1..8 come from this screen only while Write enable is ON (refused while ENABLE is active on VTDManualTest). Otherwise the PO come from VTDManualTest.'
  2187 = 'Rdy'
  2006 = 'Ready'
  2192 = 'Ready for task'
  2027 = 'REFERENCE - 300'
  2010 = 'Referenced'
  2220 = 'REQUEST ACCESS'
  2221 = 'Request only: the door is unlocked by the safety system.'
  2058 = 'RESET'
  2059 = 'RESET = drive fault reset (PO 1.8)'
  2081 = 'RESET ALL'
  2086 = 'Roller 1'
  2087 = 'Roller 2'
  2088 = 'Roller 3'
  2089 = 'Roller 4'
  2090 = 'Roller 5'
  2212 = 'ROTATE CCW'
  2213 = 'ROTATE CW'
  2098 = 'Run'
  2045 = 'RUN +'
  2044 = 'RUN -'
  2111 = 'Running'
  2130 = 'S'
  2219 = 'Safe to restart'
  2077 = 'Safety OK'
  2074 = 'SAFETY RESET'
  1086 = 'Scaling from MOVISUITE'
  2190 = 'Select a device to see the details and operate it.'
  2191 = 'Selected device'
  1060 = 'Sent'
  2049 = 'sent'
  2145 = 'Setpoint'
  1066 = 'Setpoint accel.'
  1072 = 'Setpoint appl. mode'
  1068 = 'Setpoint decel.'
  1064 = 'Setpoint speed'
  2067 = 'Settings OK'
  2233 = 'Shuttle data is not available in the PLC yet.'
  2195 = 'Shuttle high'
  2120 = 'SHUTTLES'
  2231 = 'Shuttles'
  2232 = 'SHUTTLES - screen in preparation'
  2154 = 'Signals'
  2159 = 'Slack 1'
  2160 = 'Slack 2'
  2165 = 'Slack 3'
  2166 = 'Slack 4'
  2056 = 'SOFTWARE STOP'
  2016 = 'Speed'
  2188 = 'Speed %'
  2026 = 'SPEED - 200'
  2198 = 'Speed act.'
  2197 = 'Speed req.'
  1083 = 'Speed, ramps and position in user units (scaling from MOVISUITE).'
  2048 = 'START'
  2189 = 'State'
  2136 = 'State machine'
  2125 = 'Status'
  1018 = 'Status word'
  1078 = 'Status word (PI 1)'
  1023 = 'Status/main fault - subfault'
  2005 = 'STO inactive (safety circuit OK)'
  2167 = 'STOP'
  2051 = 'STOP (normal ramp)'
  2127 = 'Stopped'
  2234 = 'System status'
  2047 = 'Target'
  1074 = 'Target pos. high'
  1076 = 'Target pos. low'
  2050 = 'Target: 400 = absolute position, 401 = relative distance. 300 = referencing.'
  1059 = 'Test'
  1111 = 'test\t'
  1080 = 'TEST ONLY - Process outputs (PLC -> drive)'
  2003 = 'TEST ONLY - SOFTWARE STOP is not an emergency stop: keep the hardwired E-stop within reach. + = positive motor direction (check up / down at the first jog).'
  2061 = 'Test settings (persistent, MOVISUITE user units)'
  1056 = 'Test write active'
  1057 = 'Timeout expired - toggle Write enable'
  2200 = 'To ID'
  1025 = 'Torque'
  2017 = 'Torque (0.1 %)'
  1084 = 'Torque PI 4 in 0.1 % of nominal motor torque.'
  2168 = 'Tower'
  2092 = 'Turntable'
  2158 = 'Ult. creep'
  2157 = 'Ult. slow'
  2170 = 'Upper limit'
  2039 = 'user units'
  2146 = 'Velocity'
  2096 = 'VTD'
  1006 = 'VTD MOVIPRO - Process Data Test (TEST ONLY)'
  2013 = 'Warning'
  1009 = 'WcState error'
  1013 = 'Word'
  327 = 'Write enable'
END_TEXTLIST

// ---- TL_Test.TcTLO
TEXTLIST TL_Test
  0 = 'Manual'
  1 = 'Semi-Auto'
  2 = 'Automatic'
   = ''
END_TEXTLIST

// ---- VISUs/Access_Gates.TcVIS
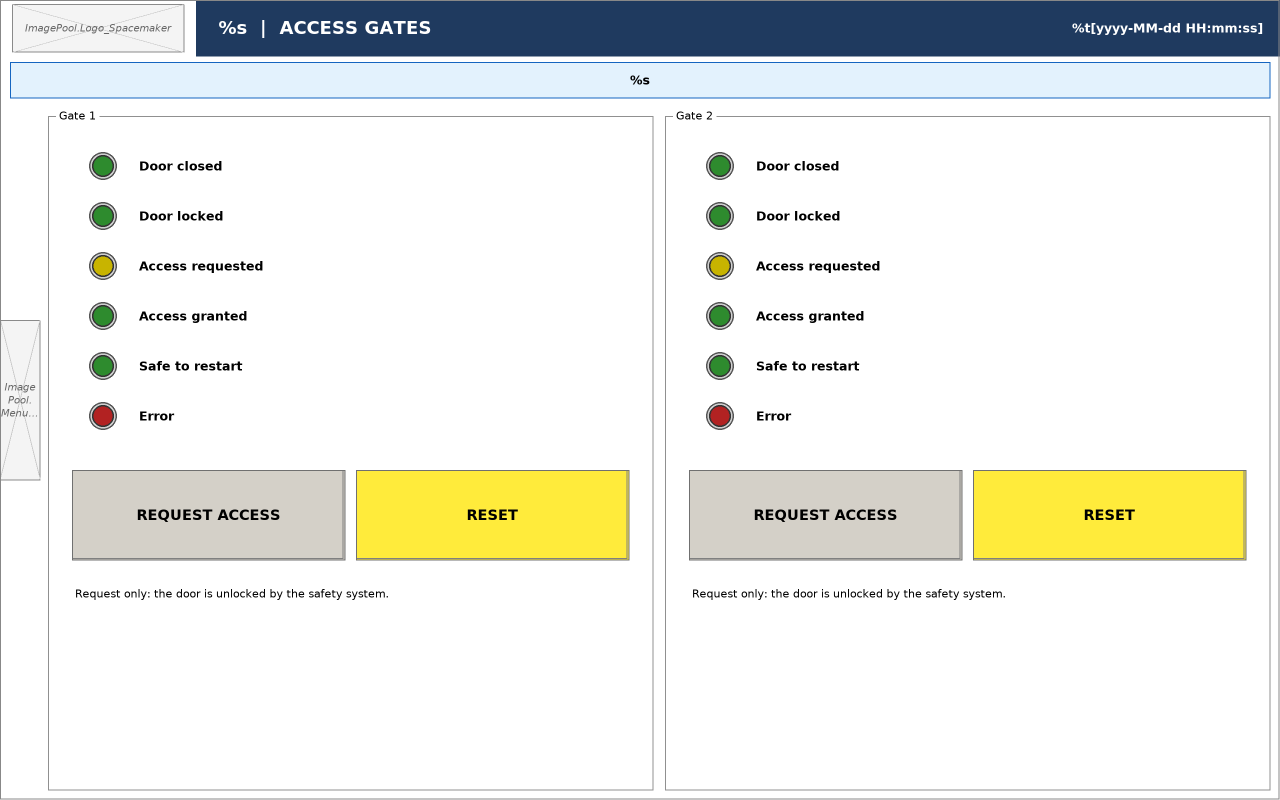
VISUALIZATION Access_Gates  // 1280x800
    Rectangle (0,0 196x56)
        OnMouseClick: change screen: Main
    Image (12,4 172x48), image: ImagePool.Logo_Spacemaker
        OnMouseClick: change screen: Main
    Rectangle (196,0 1084x56), "%s | ACCESS GATES", text variable: GVL_HMI_System.stStatus.sSystemName
    Rectangle (930,8 336x40), "%t[yyyy-MM-dd HH:mm:ss]", text variable: GVL_HMI_System.stStatus.dtNow
    Rectangle (10,62 1260x36), "%s", text variable: GVL_HMI_System.stStatus.sMessage, colour toggle: GVL_HMI_System.stStatus.bMessageAlarm
    GroupBox (48,108 605x682), "Gate 1"
    Lamp1 (87,150 32x32), variable: GVL_HMI_Gates.astGate[1].bClosed, style: Lamp-Lamp1-Green
    Rectangle (136,150 356x32), "Door closed"
    Lamp1 (87,200 32x32), variable: GVL_HMI_Gates.astGate[1].bLocked, style: Lamp-Lamp1-Green
    Rectangle (136,200 356x32), "Door locked"
    Lamp1 (87,250 32x32), variable: GVL_HMI_Gates.astGate[1].bAccessRequested, style: Lamp-Lamp1-Yellow
    Rectangle (136,250 356x32), "Access requested"
    Lamp1 (87,300 32x32), variable: GVL_HMI_Gates.astGate[1].bAccessGranted, style: Lamp-Lamp1-Green
    Rectangle (136,300 356x32), "Access granted"
    Lamp1 (87,350 32x32), variable: GVL_HMI_Gates.astGate[1].bSafeToRestart, style: Lamp-Lamp1-Green
    Rectangle (136,350 356x32), "Safe to restart"
    Lamp1 (87,400 32x32), variable: GVL_HMI_Gates.astGate[1].bError, style: Lamp-Lamp1-Red
    Rectangle (136,400 356x32), "Error"
    Button (72,470 273x90), "REQUEST ACCESS"
        tap GVL_HMI_Gates.astCommand[1].bRequestAccess p3779583253=TRUE
    Button (356,470 273x90), "RESET"
        tap GVL_HMI_Gates.astCommand[1].bReset p3779583253=TRUE
    Rectangle (72,580 557x28), "Request only: the door is unlocked by the safety system."
    GroupBox (665,108 605x682), "Gate 2"
    Lamp1 (704,150 32x32), variable: GVL_HMI_Gates.astGate[2].bClosed, style: Lamp-Lamp1-Green
    Rectangle (753,150 356x32), "Door closed"
    Lamp1 (704,200 32x32), variable: GVL_HMI_Gates.astGate[2].bLocked, style: Lamp-Lamp1-Green
    Rectangle (753,200 356x32), "Door locked"
    Lamp1 (704,250 32x32), variable: GVL_HMI_Gates.astGate[2].bAccessRequested, style: Lamp-Lamp1-Yellow
    Rectangle (753,250 356x32), "Access requested"
    Lamp1 (704,300 32x32), variable: GVL_HMI_Gates.astGate[2].bAccessGranted, style: Lamp-Lamp1-Green
    Rectangle (753,300 356x32), "Access granted"
    Lamp1 (704,350 32x32), variable: GVL_HMI_Gates.astGate[2].bSafeToRestart, style: Lamp-Lamp1-Green
    Rectangle (753,350 356x32), "Safe to restart"
    Lamp1 (704,400 32x32), variable: GVL_HMI_Gates.astGate[2].bError, style: Lamp-Lamp1-Red
    Rectangle (753,400 356x32), "Error"
    Button (689,470 273x90), "REQUEST ACCESS"
        tap GVL_HMI_Gates.astCommand[2].bRequestAccess p3779583253=TRUE
    Button (973,470 273x90), "RESET"
        tap GVL_HMI_Gates.astCommand[2].bReset p3779583253=TRUE
    Rectangle (689,580 557x28), "Request only: the door is unlocked by the safety system."
    Rectangle (0,320 40x160)
        OnMouseClick: OpenDialog Dialog=Dialog, OpenModal=True, PositionX=0, PositionY=0
        OnMouseEnter: OpenDialog Dialog=Dialog, OpenModal=True, PositionX=0, PositionY=0
    Image (0,320 40x160), image: ImagePool.Menu_Tab
        OnMouseClick: OpenDialog Dialog=Dialog, OpenModal=True, PositionX=0, PositionY=0
        OnMouseEnter: OpenDialog Dialog=Dialog, OpenModal=True, PositionX=0, PositionY=0
END_VISUALIZATION

// ---- VISUs/Alarms.TcVIS
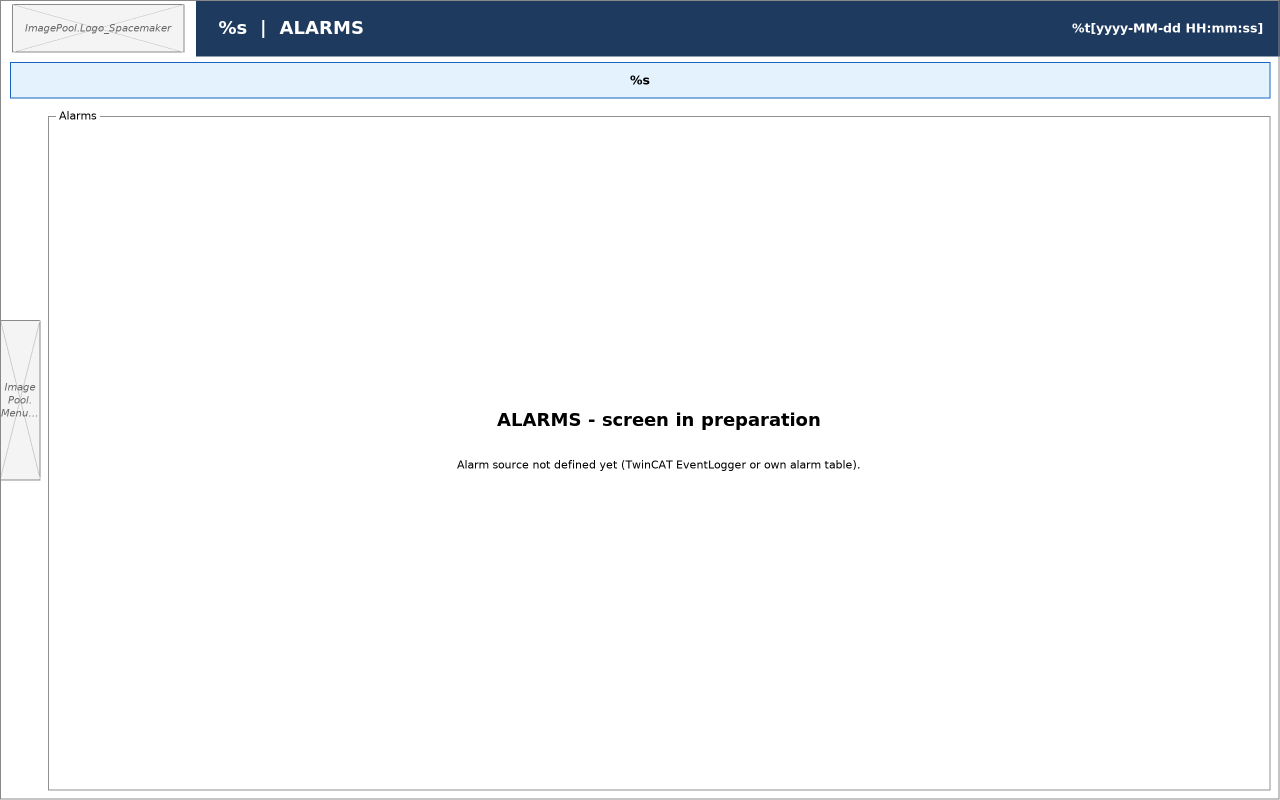
VISUALIZATION Alarms  // 1280x800
    Rectangle (0,0 196x56)
        OnMouseClick: change screen: Main
    Image (12,4 172x48), image: ImagePool.Logo_Spacemaker
        OnMouseClick: change screen: Main
    Rectangle (196,0 1084x56), "%s | ALARMS", text variable: GVL_HMI_System.stStatus.sSystemName
    Rectangle (930,8 336x40), "%t[yyyy-MM-dd HH:mm:ss]", text variable: GVL_HMI_System.stStatus.dtNow
    Rectangle (10,62 1260x36), "%s", text variable: GVL_HMI_System.stStatus.sMessage, colour toggle: GVL_HMI_System.stStatus.bMessageAlarm
    GroupBox (48,108 1222x682), "Alarms"
    Rectangle (78,400 1162x40), "ALARMS - screen in preparation"
    Rectangle (78,450 1162x30), "Alarm source not defined yet (TwinCAT EventLogger or own alarm table)."
    Rectangle (0,320 40x160)
        OnMouseClick: OpenDialog Dialog=Dialog, OpenModal=True, PositionX=0, PositionY=0
        OnMouseEnter: OpenDialog Dialog=Dialog, OpenModal=True, PositionX=0, PositionY=0
    Image (0,320 40x160), image: ImagePool.Menu_Tab
        OnMouseClick: OpenDialog Dialog=Dialog, OpenModal=True, PositionX=0, PositionY=0
        OnMouseEnter: OpenDialog Dialog=Dialog, OpenModal=True, PositionX=0, PositionY=0
END_VISUALIZATION

